(* IEC 61131-3 sources: daoli-st-library/DL_Process (part 49) *)

(* ---- FB_DL_RoMembraneFlushSeq.st ---- *)
(*
  Name: FB_DL_RoMembraneFlushSeq
  Category: DL_Process
  Version: 1.0.0
  Round: R90 / 2026-11-25
  开源溯源：clean-room 自研（族 RO/NF 膜法水处理，ST 开源生态实测 0 命中，无外部代码引入）
  功能：1) RO 停机冲洗序状态机，五相推进：待机 → 低压冲洗 → 浸泡 → 排放 → 完成。
           待机相等待 xStart 上升沿（必须边沿，防止上电即在启动位自动启动）；
           低压冲洗相开冲洗阀与浓水阀，按 tFlushS 定时并以冲洗流量监督为前置放行条件；
           浸泡相全阀关闭让药液/水在膜面停留 tSoakS；排放相只开浓水阀排空残液 DL_DRAIN_S；
           完成相置 xDone 并保持，直到 xStart 撤下才回待机（为下一次冲洗重新武装边沿）。
        2) 每相独立超时 + 整序总超时：相定时器给出正常推进点，相超时定时器给出
           「定时 + DL_OVER_MARGIN」的越限点，整序总超时由 tonTotal 兜底，
           三者并发监视，任一命中立即进故障相并锁存码值。
        3) 低液位双语义：待机相低液位只拦启动并置信息级码（不置故障位，允许液位恢复后直接启动）；
           冲洗过程中低液位判故障（泵空转保护）。
  边界条件：1) 非有限值闸：冲洗流量入参过 NOT(x > -DL_BIG AND x < DL_BIG)，同时拦 NaN 与 Inf；
           命中即判流量监督不通过（_bFlowOk := FALSE），由流量宽限定时器升级为故障，
           绝不把 NaN 直接与 DL_FLOW_MIN 比较（NaN 比较恒假会伪装成「流量正常」，R19）。
        2) 时间参数零闸：tFlushS / tSoakS <= T#0S 时对应相定时器立即置 Q，等价于该相跳过；
           这是合法组态（调试用），不判无效，但语义在此声明，禁止下游按「必有停留」假设。
        3) 流量下限零闸：DL_FLOW_MIN > DL_EPS，且流量监督只在低压冲洗相生效（其余相无流量要求）。
        4) 饱和与钳制：冲洗流量不做数值钳制（只做比较，不参与运算），避免掩盖超量程故障；
           所有相迁移均以定时器 Q 位与状态量为门控，不以单拍布尔标志门控（R274）。
        5) 故障解除路径：故障相内 (NOT xStart) AND (NOT xFault) 成立即清锁存回待机；
           回待机后必须重新给 xStart 上升沿才能再启动（rtStart 已被清，不会自恢复）。
        6) 状态机兜底：CASE 全态覆盖 + ELSE 强制回故障相并清全部输出。
        7) FB 主体不使用 RETURN，统一单出口（跨平台可移植性）。
  量纲自证：fFlushFlowM3h 为体积流量 [m3/h]，仅与同量纲的 DL_FLOW_MIN [m3/h] 比较；
           tFlushS / tSoakS / DL_DRAIN_S / DL_OVER_MARGIN / DL_TOTAL_MAX 全部为 [TIME]，
           相超时点 = [TIME] + [TIME] = [TIME]，与 TON 的 PT 同量纲；
           本件不出现跨量纲相加（无功率/温度/压力混合运算）。
  码表 Error codes（本件格 0090_03xx，故障级一律 3 行内置 _uFault/_bFault/_eState）:
    16#0090_0301 信息级：低液位，禁止启动冲洗（不置故障位）
    16#0090_0302 故障级：低压冲洗相冲洗流量不足（宽限窗超时）
    16#0090_0303 故障级：低压冲洗相超时（定时已到但放行条件不满足）
    16#0090_0304 故障级：浸泡相超时
    16#0090_0305 故障级：排放相超时
    16#0090_0306 故障级：整序总超时
    16#0090_0307 故障级：外部故障输入 xFault
    16#0090_0308 故障级：冲洗过程中低液位（泵空转保护）
    16#0090_0309 故障级：状态机落 ELSE 兜底（非法相位 ID）

  修订历史 Revision :
    2026-11-25  v1.0.0  R90 首版
*)

TYPE E_DL_RoFlushState :
(
    eRoFlushIdle     := 0,    // 待机：等启动上升沿 / Idle, awaiting start rising edge
    eRoFlushLowPress := 10,   // 低压冲洗：冲洗阀 + 浓水阀开 / Low-pressure flush, both valves open
    eRoFlushSoak     := 20,   // 浸泡：全阀关闭保持 / Soak, all valves closed
    eRoFlushDrain    := 30,   // 排放：仅浓水阀开排空 / Drain, concentrate valve only
    eRoFlushDone     := 40,   // 完成：xDone 保持至撤令 / Done, held until start released
    eRoFlushFault    := 90    // 故障：锁存待解除 / Fault, latched awaiting release
);
END_TYPE

FUNCTION_BLOCK FB_DL_RoMembraneFlushSeq
VAR_INPUT
    xStart        : BOOL;    // 冲洗启动指令（上升沿有效）[bool] / Flush start command, edge triggered [bool]
    xFault        : BOOL;    // 外部故障汇总 [bool] / External fault aggregate [bool]
    xLowLevel     : BOOL;    // 水箱低液位开关 [bool] / Tank low level switch [bool]
    fFlushFlowM3h : REAL;    // 冲洗水实测体积流量 [m3/h] / Measured flush water flow [m3/h]
    tFlushS       : TIME;    // 低压冲洗设定时长 [TIME] / Low-pressure flush duration [TIME]
    tSoakS        : TIME;    // 浸泡设定时长 [TIME] / Soak duration [TIME]
END_VAR
VAR_OUTPUT
    xFlushValve   : BOOL;    // 冲洗进水阀指令（安全侧：故障时关）[bool] / Flush inlet valve command [bool]
    xBrineValve   : BOOL;    // 浓水排放阀指令（安全侧：故障时关）[bool] / Brine discharge valve command [bool]
    xDone         : BOOL;    // 冲洗完成保持位 [bool] / Flush complete held flag [bool]
    xBusy         : BOOL;    // 冲洗进行中 [bool] / Flush sequence busy [bool]
    xFlowOk       : BOOL;    // 冲洗流量监督通过 [bool] / Flush flow supervision passed [bool]
    eState        : E_DL_RoFlushState;   // 状态出口，段尾单点映射 / State outlet, single-point mapped
    nErrId        : UDINT;   // 事件码，0 = 无事件 / Event code, 0 = none
END_VAR
VAR
    tonFlush      : TON;     // 低压冲洗相正常定时 [TIME] / Low-pressure flush phase timer
    tonFlushOv    : TON;     // 低压冲洗相超时定时 [TIME] / Low-pressure flush overrun timer
    tonSoak       : TON;     // 浸泡相正常定时 [TIME] / Soak phase timer
    tonSoakOv     : TON;     // 浸泡相超时定时 [TIME] / Soak overrun timer
    tonDrain      : TON;     // 排放相正常定时 [TIME] / Drain phase timer
    tonDrainOv    : TON;     // 排放相超时定时 [TIME] / Drain overrun timer
    tonTotal      : TON;     // 整序总超时定时 [TIME] / Whole-sequence total timeout timer
    tonFlowG      : TON;     // 冲洗流量宽限定时 [TIME] / Flush flow grace timer
    rtStart       : R_TRIG;  // 启动上升沿检测 [bool] / Start rising edge detector
    _eState       : E_DL_RoFlushState := E_DL_RoFlushState.eRoFlushIdle;   // 内部相位（CASE 唯一写入目标）
    _eStatePrev   : E_DL_RoFlushState := E_DL_RoFlushState.eRoFlushIdle;   // 上一拍相位快照（周期末更新）
    _bFlowOk      : BOOL;    // 冲洗流量监督结果 [bool] / Flush flow supervision result [bool]
    _bActive      : BOOL;    // 序激活（三执行相之一）[bool] / Sequence active flag [bool]
    _bDoneL       : BOOL;    // 完成位锁存（跨相保持）[bool] / Done latch held across phases [bool]
    _bFault       : BOOL;    // 故障锁存位 [bool] / Latched fault flag [bool]
    _uInfo        : UDINT;   // 信息码，每拍重算 / Info code, recomputed every cycle
    _uFault       : UDINT;   // 故障码锁存 / Latched fault code
    _iPhaseChg    : INT;     // 本拍相位切换计数（观测用）[-] / Phase-change count this cycle [-]
END_VAR
VAR CONSTANT
    DL_EPS        : REAL := 1.0E-9;      // 数值零闸阈值 [-] / Numeric zero gate threshold [-]
    DL_BIG        : REAL := 1.0E12;      // 非有限值闸量级上限 [-] / Finiteness gate magnitude [-]
    DL_FLOW_MIN   : REAL := 0.50;        // 冲洗流量监督下限 [m3/h] / Flush flow supervision low [m3/h]
    DL_DRAIN_S    : TIME := T#20S;       // 排放相设定时长 [TIME] / Drain phase duration [TIME]
    DL_OVER_MARGIN: TIME := T#30S;       // 相超时相对正常定时的裕量 [TIME] / Phase overrun margin [TIME]
    DL_TOTAL_MAX  : TIME := T#2H;        // 整序总超时上限 [TIME] / Whole-sequence total timeout [TIME]
    DL_FLOW_GRACE : TIME := T#10S;       // 冲洗流量不足宽限窗 [TIME] / Flow-shortage grace window [TIME]
END_VAR

(* —— 段 0：单拍量预清零（锁存量 _uFault/_bFault/_bDoneL/_eStatePrev 不入清单，R187①） —— *)
_uInfo := 16#0000_0000;                     // 信息码每拍重算 / Info code recomputed
_iPhaseChg := 0;                            // 相位切换计数每拍重算 / Phase-change counter recomputed
nErrId := 16#0000_0000;                     // 事件码缺省无事件 / Event code defaults to none

(* —— 段 1：非有限值闸（R19：流量不参与运算，但必须拦住 NaN 比较的伪装成真） —— *)
IF NOT (fFlushFlowM3h > -DL_BIG AND fFlushFlowM3h < DL_BIG) THEN
    _bFlowOk := FALSE;                      // 非有限一律判流量不通过（不是运算符，是安全侧）
ELSE
    _bFlowOk := (fFlushFlowM3h >= DL_FLOW_MIN);   // 与同量纲下限比较 [m3/h] vs [m3/h]
END_IF

(* —— 段 2：状态派生量（本拍相位为上一拍末值，标准 FB 周期语义） —— *)
_bActive := (_eState = E_DL_RoFlushState.eRoFlushLowPress)
            OR (_eState = E_DL_RoFlushState.eRoFlushSoak)
            OR (_eState = E_DL_RoFlushState.eRoFlushDrain);

(* —— 段 3：定时器与边沿无条件周期刷新（R7：调用语句不得置于 IF/CASE 内） —— *)
rtStart(CLK := xStart);                                                      // 启动上升沿，每拍必调
tonFlush(IN := (_eState = E_DL_RoFlushState.eRoFlushLowPress), PT := tFlushS);            // 冲洗相正常定时
tonFlushOv(IN := (_eState = E_DL_RoFlushState.eRoFlushLowPress),
           PT := tFlushS + DL_OVER_MARGIN);                                  // 冲洗相超时点 = 定时 + 裕量
tonSoak(IN := (_eState = E_DL_RoFlushState.eRoFlushSoak), PT := tSoakS);                  // 浸泡相正常定时
tonSoakOv(IN := (_eState = E_DL_RoFlushState.eRoFlushSoak),
          PT := tSoakS + DL_OVER_MARGIN);                                    // 浸泡相超时点
tonDrain(IN := (_eState = E_DL_RoFlushState.eRoFlushDrain), PT := DL_DRAIN_S);            // 排放相正常定时
tonDrainOv(IN := (_eState = E_DL_RoFlushState.eRoFlushDrain),
           PT := DL_DRAIN_S + DL_OVER_MARGIN);                               // 排放相超时点
tonTotal(IN := _bActive, PT := DL_TOTAL_MAX);                                // 整序总超时，自复位由相位驱动
tonFlowG(IN := (_eState = E_DL_RoFlushState.eRoFlushLowPress) AND (NOT _bFlowOk),
         PT := DL_FLOW_GRACE);                                               // 流量不足宽限窗

(* —— 段 4：全局故障拦截（优先级最高；已锁存则不再改写码值，禁同拍抹除） —— *)
IF xFault AND (NOT _bFault) THEN
    _uFault := 16#0090_0307;                // 故障级：外部故障输入
    _bFault := TRUE;                        // 锁存（3 行内置，R45 配对）
    _eState := E_DL_RoFlushState.eRoFlushFault;
END_IF
IF tonTotal.Q AND _bActive AND (NOT _bFault) THEN
    _uFault := 16#0090_0306;                // 故障级：整序总超时
    _bFault := TRUE;                        // 锁存
    _eState := E_DL_RoFlushState.eRoFlushFault;
END_IF

(* —— 段 5：相位机（只做迁移；出口在段 7 单点映射） —— *)
CASE _eState OF

E_DL_RoFlushState.eRoFlushIdle:
    IF NOT xStart THEN
        _bDoneL := FALSE;                   // 撤令即清完成位，为下次冲洗重新武装
    ELSIF xLowLevel THEN
        _uInfo := 16#0090_0301;             // 信息级：低液位禁止启动（不置故障位）
    ELSIF rtStart.Q THEN
        _bDoneL := FALSE;                   // 新序开始：清完成位（迁移前一次性清）
        _eState := E_DL_RoFlushState.eRoFlushLowPress;   // 进低压冲洗相
    END_IF

E_DL_RoFlushState.eRoFlushLowPress:
    IF xLowLevel THEN
        _uFault := 16#0090_0308;            // 故障级：冲洗中低液位（泵空转保护）
        _bFault := TRUE;
        _eState := E_DL_RoFlushState.eRoFlushFault;
    ELSIF tonFlush.Q AND _bFlowOk THEN
        _eState := E_DL_RoFlushState.eRoFlushSoak;       // 本拍合法事件优先于超时迁移（R275）
    ELSIF tonFlowG.Q THEN
        _uFault := 16#0090_0302;            // 故障级：冲洗流量不足
        _bFault := TRUE;
        _eState := E_DL_RoFlushState.eRoFlushFault;
    ELSIF tonFlushOv.Q THEN
        _uFault := 16#0090_0303;            // 故障级：低压冲洗相超时
        _bFault := TRUE;
        _eState := E_DL_RoFlushState.eRoFlushFault;
    END_IF

E_DL_RoFlushState.eRoFlushSoak:
    IF xLowLevel THEN
        _uFault := 16#0090_0308;            // 故障级：浸泡中低液位
        _bFault := TRUE;
        _eState := E_DL_RoFlushState.eRoFlushFault;
    ELSIF tonSoak.Q THEN
        _eState := E_DL_RoFlushState.eRoFlushDrain;      // 浸泡到点：进排放相
    ELSIF tonSoakOv.Q THEN
        _uFault := 16#0090_0304;            // 故障级：浸泡相超时
        _bFault := TRUE;
        _eState := E_DL_RoFlushState.eRoFlushFault;
    END_IF

E_DL_RoFlushState.eRoFlushDrain:
    IF xLowLevel THEN
        _uFault := 16#0090_0308;            // 故障级：排放中低液位
        _bFault := TRUE;
        _eState := E_DL_RoFlushState.eRoFlushFault;
    ELSIF tonDrain.Q THEN
        _bDoneL := TRUE;                    // 完成位锁存（跨相保持，段 7 单点映射）
        _eState := E_DL_RoFlushState.eRoFlushDone;       // 进完成相
    ELSIF tonDrainOv.Q THEN
        _uFault := 16#0090_0305;            // 故障级：排放相超时
        _bFault := TRUE;
        _eState := E_DL_RoFlushState.eRoFlushFault;
    END_IF

E_DL_RoFlushState.eRoFlushDone:
    IF xFault THEN
        _uFault := 16#0090_0307;            // 故障级：完成后外部故障（段 4 已拦，此处兜底同码）
        _bFault := TRUE;
        _eState := E_DL_RoFlushState.eRoFlushFault;
    ELSIF NOT xStart THEN
        _bDoneL := FALSE;                   // 撤令：清完成位并回待机
        _eState := E_DL_RoFlushState.eRoFlushIdle;
    END_IF

E_DL_RoFlushState.eRoFlushFault:
    IF (NOT xStart) AND (NOT xFault) THEN
        _bFault := FALSE;                   // 解除路径：撤令 AND 外部故障消失（可达）
        _uFault := 16#0000_0000;            // 清锁存码
        _bDoneL := FALSE;                   // 完成位一并清，避免故障后误报完成
        _eState := E_DL_RoFlushState.eRoFlushIdle;       // 回待机，需新上升沿才可再启动
    END_IF

ELSE
    _uFault := 16#0090_0309;                // 故障级：非法相位 ID 兜底
    _bFault := TRUE;                        // 锁存
    _eState := E_DL_RoFlushState.eRoFlushFault;          // 强制回故障相

END_CASE

(* —— 段 6：后置段（R23：相位切换后的清计数与快照统一放在迁移判断之后） —— *)
IF _eState <> _eStatePrev THEN
    _iPhaseChg := _iPhaseChg + 1;           // 相位已切换：记一拍切换事件（观测用）
END_IF
_eStatePrev := _eState;                     // 快照在周期末尾统一更新，禁跨相重试预算不清零

(* —— 段 7：出口单点映射（名实同源；阀门由状态导出，不在多分支各写一遍，故障侧一律关） —— *)
xFlushValve := (_eState = E_DL_RoFlushState.eRoFlushLowPress) AND (NOT _bFault);      // 仅冲洗相开
xBrineValve := ((_eState = E_DL_RoFlushState.eRoFlushLowPress)
                OR (_eState = E_DL_RoFlushState.eRoFlushDrain)) AND (NOT _bFault);    // 冲洗/排放相开
xDone := _bDoneL AND (NOT _bFault);                                                      // 完成位出口
xBusy := _bActive AND (NOT _bFault);                                                     // 进行中出口
xFlowOk := _bFlowOk;                                                                     // 流量监督出口
eState := _eState;                                                                       // 状态出口单点映射
IF _bFault THEN
    nErrId := _uFault;                      // 故障锁存码回放（不在故障相按当下输入重推断）
ELSE
    nErrId := _uInfo;                       // 信息码
END_IF

END_FUNCTION_BLOCK

(* ---- FB_DL_RoomClimateCtrl.st ---- *)
//==============================================================================
// 功能块：FB_DL_RoomClimateCtrl ｜ 中文名称：房间温湿度双回路耦合控制
// 所属子库：DL_Process ｜ 版本：v1.0.1 ｜ 兼容：CODESYS V3.5+ / TwinCAT 3 / 汇川 InoProShop
// 功能描述：房间温湿度双回路耦合控制：温度回路单 PID 带符号输出分程
//           （正 = 加热阀、负 = 冷却阀），湿度回路单 PID 带符号输出分
//           程（正 = 加湿阀、负 = 除湿阀），带宽死区内输出保持（PID
//           内置死区）。防结露联锁（安全联锁而非优化，头注释写明物理
//           后果：供水温度低于「露点 + 余量」时冷盘管表面结露滴水，
//           滴水进入洁净室即污染事故）→ 限制冷却/除湿阀上限并置
//           bCondensationRisk + 信息 0401。温湿同拍冲突互斥仲裁（冷侧
//           优先：冷却与加湿同拍 → 撤加湿；除湿与加热同拍 → 撤加热，
//           均置 bConflictArbitrated + 信息 0400）。PID 组合调用
//           FB_DL_PidController（两实例，不内联），露点由
//           FC_DL_DewPointCalc 计算（Magnus-Tetens 常数唯一属主
//           FC_DL_VaporPressureSat，R23 裁定，只调用不复制）。失能四
//           阀回 0%（安全侧：不制冷不加热不加湿不除湿）。
// 开源溯源 (Origin)：道莅 clean-room 防御性实现（仅借 OSCAT ROOM_CONTROL 行为定义/参数域，零代码行与符号名复制）
// 单位表：温度[摄氏度] / 相对湿度[%] / 带宽[K 或百分数] / 阀输出[百分数] / 增益[百分数每K 或 百分数每百分数] / 积分时间[s] / 余量[K] / 扫描间隔[ms]
// 错误码表：16#0005_0400 信息级（温湿回路同拍冲突被互斥仲裁，冷侧优先，
//           不置 bError）/ 16#0005_0401 信息级（防结露联锁限制降温与
//           除湿，安全联锁生效，不置 bError）/ 16#0005_0342 故障级（设
//           定域/带宽/增益/余量组态非法，置 bError）/ 16#0005_0343 故
//           障级（输入非有限，置 bError，四阀回 0% 安全侧）/
//           16#0005_0344 故障级兜底（状态机落 ELSE 或非法状态，置
//           bError 并四阀回 0%）
// 状态机：E_DL_RoomClimateState（eIdle=0 / eAuto=10 / eInterlock=20 /
//           eFault=99），CASE 含 ELSE 兜底，ELSE 置 0344 并四阀回 0%
//           （安全侧：联锁与仲裁之外任何异常一律全关执行器）
// 边界行为：① 冷/热阀互斥（分程结构天然互斥），跨回路同拍冲突仲裁：
//           冷侧优先（冷却 ∧ 加湿 → 撤加湿；除湿 ∧ 加热 → 撤加热），
//           置 bConflictArbitrated + 信息 0400；② 防结露联锁：
//           fChwSupplyC 低于露点 + fDewMarginK → bCondensationRisk +
//           信息 0401，冷却/除湿阀上限按 (供水 − 露点)/余量 线性压缩
//           （供水贴露点 → 0%，供水达露点 + 余量 → 100%），这是安全
//           联锁而非优化；③ 带宽死区内 PID 输出保持（防阀频繁动作）；
//           ④ 设定域/带宽/增益/余量组态非法（带宽非正、温度设定超
//           0~45、湿度设定超 10~95、增益非正、余量小于 0）→ 故障 0342；
//           ⑤ 非有限（NaN 自反判 + Inf 幅值上限判，R79）→ 故障 0343，
//           四阀回 0% 安全侧；⑥ 失能 → 四阀回 0% + bValid := FALSE
//           （安全侧：不制冷不加热不加湿不除湿）；⑦ 双 PID 与露点件
//           每拍无条件调用恰好一次（实例纪律）；⑧ 贴限 bAtLimit：任
//           一阀达 100%（容差比较）；⑨ 上电首拍 bValid := FALSE。
// 修订历史：v1.0.0 2026-11-17 首版（R25 派单 · §4.10，依赖 §4.1 件语义）
//           v1.0.1 2026-11-17 终审补失能出口收口（段 11，对外引脚契约零变更）：PID 件失能时
//           输出回 rOutMin = −100%，经带符号分程映射为 100% 冷却/除湿，而四阀归零只在下一拍
//           eIdle 相执行，导致「失能 = 四阀回 0%」契约在失能沿那一拍被破坏（安全侧漂移）。
//           收口放在 CASE 之后：失能电平期间出口强制 0%（不依赖相切换时序）。
//==============================================================================
(*------------------------------------------------------------------------------
 * 枚举: E_DL_RoomClimateState（归属 DL_Process，与 FB_DL_RoomClimateCtrl 同文件）
 *----------------------------------------------------------------------------*)
TYPE E_DL_RoomClimateState :
(
    eIdle      := 0,   // 失能/待机：四阀回 0% / Idle: all four valves closed
    eAuto      := 10,  // 双回路自动：分程输出无联锁限制 / Auto: split-range outputs, no interlock
    eInterlock := 20,  // 防结露联锁生效：冷却/除湿被限幅 / Anti-condensation interlock: cooling and dehumidifying capped
    eFault     := 99   // 故障兜底态：组态非法/非有限/非法状态，四阀回 0% / Fault fallback, valves closed
);
END_TYPE
FUNCTION_BLOCK FB_DL_RoomClimateCtrl
VAR_INPUT
    fTempSetC      : LREAL;                    // 温度设定 [摄氏度]，域 0~45 / Temperature setpoint [degC], domain 0..45
    fTempMeasC     : LREAL;                    // 实测温度 [摄氏度] / Measured temperature [degC]
    fRhSetPct      : LREAL;                    // 湿度设定 [百分数]，域 10~95 / Humidity setpoint [percent], domain 10..95
    fRhMeasPct     : LREAL;                    // 实测湿度 [百分数] / Measured humidity [percent]
    fTempBandK     : LREAL := 0.5;             // 温度带宽 [K]，死区内输出保持 / Temperature dead band [K]
    fRhBandPct     : LREAL := 3.0;             // 湿度带宽 [百分数] / Humidity dead band [percent]
    fChwSupplyC    : LREAL;                    // 冷冻水供水温度 [摄氏度]，防结露用 / Chilled-water supply temperature [degC]
    fDewMarginK    : LREAL := 1.5;             // 防结露安全余量 [K] / Anti-condensation margin [K]
    fKpValvePctPerK : LREAL := 12.0;           // 温度回路比例增益 [百分数每K] / Temperature loop proportional gain [percent per K]
    fTiTempS       : LREAL := 180.0;           // 温度回路积分时间 [s]，0 = 纯比例 / Temperature loop integral time [s]
    fKpDehumPctPerPct : LREAL := 5.0;          // 湿度回路比例增益 [百分数每百分数] / Humidity loop proportional gain [percent per percent]
    fTiRhS         : LREAL := 240.0;           // 湿度回路积分时间 [s]，0 = 纯比例 / Humidity loop integral time [s]
    uDeltaTimeMs   : UDINT;                    // 扫描间隔 [ms]，调用方注入，禁用系统时间函数 / Scan interval [ms], caller-injected
    bEnable        : BOOL;                     // 总使能 / Master enable
    bReset         : BOOL;                     // 复位，上升沿清状态与双 PID / Reset, rising edge clears state and both PIDs
END_VAR
VAR_OUTPUT
    fCoolValvePct  : LREAL;                    // 冷却阀指令 [百分数]，与加热阀互斥 / Cooling valve command [percent], exclusive with heating
    fHeatValvePct  : LREAL;                    // 加热阀指令 [百分数]，与冷却阀互斥 / Heating valve command [percent], exclusive with cooling
    fDehumValvePct : LREAL;                    // 除湿阀指令 [百分数]，与加湿阀互斥 / Dehumidifying valve command [percent], exclusive with humidifying
    fHumValvePct   : LREAL;                    // 加湿阀指令 [百分数]，与除湿阀互斥 / Humidifying valve command [percent], exclusive with dehumidifying
    bCondensationRisk : BOOL;                 // 防结露联锁生效标志 / Anti-condensation interlock active flag
    bConflictArbitrated : BOOL;                // 同拍冲突被仲裁标志（冷侧优先）/ Conflict arbitrated this scan, cold side wins
    fDewPointC     : LREAL;                    // 室内露点 [摄氏度]，下游件计算透传 / Room dew point [degC], passed through
    bAtLimit       : BOOL;                     // 任一阀达 100% / Any valve at 100 percent
    eErr           : UDINT;                    // 错误码，0 = 无错，码位 16#0005_0400 起信息级、16#0005_0342 起故障级（分带见错误码表） / Error code, 0 = no error, band info/fault per the code table
    bError         : BOOL;                     // 故障级标志，仅故障级错误置位 / Fault-class flag, set only on fault-level codes
    bValid         : BOOL;                     // 控制输出可用标志，失能/故障闸显式 FALSE / Control usable flag, explicit FALSE on disable/fault gates
    eState         : E_DL_RoomClimateState;    // 主状态机当前状态 / Current state of the main state machine
END_VAR
VAR
    fbReset        : R_TRIG;                   // 复位上升沿检测实例 / Reset rising edge detector
    fbPidTemp      : FB_DL_PidController;      // 温度回路 PID 组合实例（DL_Algo，契约见手册）/ Temperature loop PID composed instance
    fbPidRh        : FB_DL_PidController;      // 湿度回路 PID 组合实例（DL_Algo，契约见手册）/ Humidity loop PID composed instance
    fTempReal      : REAL;                     // 温度设定降精度暂存 [摄氏度] / Temperature setpoint staging in REAL precision
    fTempMeasReal  : REAL;                     // 实测温度降精度暂存 [摄氏度] / Measured temperature staging in REAL precision
    fRhSetReal     : REAL;                     // 湿度设定降精度暂存 [百分数] / Humidity setpoint staging in REAL precision
    fRhMeasReal    : REAL;                     // 实测湿度降精度暂存 [百分数] / Measured humidity staging in REAL precision
    fTempOutReal   : REAL;                     // 温度 PID 带符号输出暂存 [百分数] / Signed temperature PID output staging
    fRhOutReal     : REAL;                     // 湿度 PID 带符号输出暂存 [百分数] / Signed humidity PID output staging
    fTempSetClamped : LREAL;                   // 钳位后温度设定 [摄氏度] / Clamped temperature setpoint [degC]
    fRhSetClamped  : LREAL;                    // 钳位后湿度设定 [百分数] / Clamped humidity setpoint [percent]
    fTempRealIn    : REAL;                     // 露点件干球输入暂存 [摄氏度] / Dew-point dry-bulb staging
    fRhRealIn      : REAL;                     // 露点件湿度输入暂存 [百分数] / Dew-point humidity staging
    fDewReal       : REAL;                     // 露点返回值暂存 [摄氏度] / Dew-point return staging
    uDewErr        : UDINT;                    // 露点件错误码暂存 / Dew-point error code staging
    fVaporPa       : REAL;                     // 露点件水汽压暂存 [Pa]（诊断透传）/ Dew-point vapor pressure staging [Pa]
    bDewInRange    : BOOL;                     // 露点件域内标志暂存 / Dew-point in-domain flag staging
    bDewOk         : BOOL;                     // 露点件结果可用判据 / Dew-point usable predicate
    fCapPct        : LREAL;                    // 联锁阀位上限 [百分数] / Interlock valve cap [percent]
    fTiTempMs      : LREAL;                    // 温度回路积分时间换算毫秒 [ms] / Temperature integral time in ms
    fTiRhMs        : LREAL;                    // 湿度回路积分时间换算毫秒 [ms] / Humidity integral time in ms
    tPidSample     : TIME;                     // PID 采样周期 [ms]（扫描间隔下限钳位）/ PID sample period, floored scan interval
    ePidErr        : UDINT;                    // PID 件错误码暂存（共用判据）/ PID error code staging
    bPidErrTemp    : BOOL;                     // 温度 PID 故障标志暂存 / Temperature PID fault flag staging
    bPidErrRh      : BOOL;                     // 湿度 PID 故障标志暂存 / Humidity PID fault flag staging
    bAnyFault      : BOOL;                     // 本拍任一 PID 故障 / Any PID fault this scan
    bFirstScan     : BOOL := TRUE;             // 上电首拍标志 / First-scan flag
END_VAR
VAR CONSTANT
    DL_RCC_CODE_INFO_1 : UDINT := 16#0005_0400;   // 信息级槽 1（同拍冲突仲裁） / info slot 1
    DL_RCC_CODE_INFO_2 : UDINT := 16#0005_0401;   // 信息级槽 2（防结露联锁生效） / info slot 2
    DL_RCC_CODE_FLT_1  : UDINT := 16#0005_0342;   // 故障级槽 1（设定域/带宽组态非法） / fault slot 1
    DL_RCC_CODE_FLT_2  : UDINT := 16#0005_0343;   // 故障级槽 2（输入非有限） / fault slot 2
    DL_RCC_CODE_FLT_3  : UDINT := 16#0005_0344;   // 故障级槽 3（非法状态兜底） / fault slot 3, illegal-state fallback
    DL_RC_ZERO     : LREAL := 0.0;            // 零值常量，避免裸字面量 [—] / Zero constant, avoids a bare literal
    DL_RC_TOL      : LREAL := 1.0E-6;         // 浮点比较容差 [—] / Float comparison tolerance
    DL_RC_INF      : LREAL := 1.7976931348623157E308;  // LREAL 幅值上限，Inf 判据 / LREAL magnitude ceiling, Inf criterion
    DL_RC_TEMP_MIN : LREAL := 0.0;            // 温度设定域下限 [摄氏度] / Temperature setpoint domain floor [degC]
    DL_RC_TEMP_MAX : LREAL := 45.0;           // 温度设定域上限 [摄氏度] / Temperature setpoint domain ceiling [degC]
    DL_RC_RH_MIN   : LREAL := 10.0;           // 湿度设定域下限 [百分数] / Humidity setpoint domain floor [percent]
    DL_RC_RH_MAX   : LREAL := 95.0;           // 湿度设定域上限 [百分数] / Humidity setpoint domain ceiling [percent]
    DL_RC_T_MIN    : LREAL := -40.0;          // 露点件干球钳位下限 [摄氏度] / Dew-point dry-bulb clamp floor [degC]
    DL_RC_T_MAX    : LREAL := 60.0;           // 露点件干球钳位上限 [摄氏度] / Dew-point dry-bulb clamp ceiling [degC]
    DL_RC_RH_C_MIN : LREAL := 1.0;            // 露点件湿度钳位下限 [百分数] / Dew-point humidity clamp floor [percent]
    DL_RC_RH_C_MAX : LREAL := 100.0;          // 露点件湿度钳位上限 [百分数] / Dew-point humidity clamp ceiling [percent]
    DL_RC_OUT_MAX  : LREAL := 100.0;          // 阀输出上限 [百分数] / Valve output ceiling [percent]
    DL_RC_TD_OFF   : TIME := T#0S;            // 微分关闭语义值 [s] / Derivative-off semantic value
    DL_RC_MS_PER_S : LREAL := 1000.0;         // 毫秒转秒系数 [s/ms] / Ms-to-s factor
    DL_RC_DT_MIN_MS : UDINT := 10;            // 扫描间隔下限 [ms] / Scan interval floor [ms]
END_VAR

(*------------------------------------------------------------------------------
 * 段 1｜无条件刷新区（红线 5）：复位沿检测在任何分支之外周期调用
 *----------------------------------------------------------------------------*)
fbReset(CLK := bReset);                        // 复位沿检测无条件刷新 / reset edge refreshed unconditionally

(*------------------------------------------------------------------------------
 * 段 2｜复位沿处理（改写置于沿后，防吞沿 R39）
 *----------------------------------------------------------------------------*)
IF fbReset.Q THEN
    eState := E_DL_RoomClimateState.eIdle;
    eErr   := 16#0000_0000;                    // 复位清码 / reset clears code
    bError := FALSE;                           // 复位清故障 / reset clears fault
    bCondensationRisk := FALSE;                // 联锁标志清 / interlock flag cleared
    bConflictArbitrated := FALSE;              // 仲裁标志清 / arbitration flag cleared
    bFirstScan := TRUE;                        // 重新首拍化 / re-initialize first scan
END_IF

(*------------------------------------------------------------------------------
 * 段 3｜非有限输入闸（浮点引脚逐个：NaN 自反判 + Inf 幅值上限判，R79）
 *       命中即四阀回 0% 安全侧
 *----------------------------------------------------------------------------*)
IF (fTempSetC <> fTempSetC) OR (ABS(fTempSetC) >= DL_RC_INF)
   OR (fTempMeasC <> fTempMeasC) OR (ABS(fTempMeasC) >= DL_RC_INF)
   OR (fRhSetPct <> fRhSetPct) OR (ABS(fRhSetPct) >= DL_RC_INF)
   OR (fRhMeasPct <> fRhMeasPct) OR (ABS(fRhMeasPct) >= DL_RC_INF)
   OR (fTempBandK <> fTempBandK) OR (ABS(fTempBandK) >= DL_RC_INF)
   OR (fRhBandPct <> fRhBandPct) OR (ABS(fRhBandPct) >= DL_RC_INF)
   OR (fChwSupplyC <> fChwSupplyC) OR (ABS(fChwSupplyC) >= DL_RC_INF)
   OR (fDewMarginK <> fDewMarginK) OR (ABS(fDewMarginK) >= DL_RC_INF)
   OR (fKpValvePctPerK <> fKpValvePctPerK) OR (ABS(fKpValvePctPerK) >= DL_RC_INF)
   OR (fTiTempS <> fTiTempS) OR (ABS(fTiTempS) >= DL_RC_INF)
   OR (fKpDehumPctPerPct <> fKpDehumPctPerPct) OR (ABS(fKpDehumPctPerPct) >= DL_RC_INF)
   OR (fTiRhS <> fTiRhS) OR (ABS(fTiRhS) >= DL_RC_INF) THEN
    eState := E_DL_RoomClimateState.eFault;
    eErr   := DL_RCC_CODE_FLT_2;               // 故障级：输入非有限 / fault: non-finite input
    bError := TRUE;                            // 故障级必置 bError（R45 配对）/ fault-class pairs with bError
    bValid := FALSE;                           // 输出不可用 / outputs unusable
    fCoolValvePct := DL_RC_ZERO;               // 四阀回 0% 安全侧 / valves to zero, safe side
    fHeatValvePct := DL_RC_ZERO;               // 四阀回 0% 安全侧 / valves to zero, safe side
    fDehumValvePct := DL_RC_ZERO;              // 四阀回 0% 安全侧 / valves to zero, safe side
    fHumValvePct := DL_RC_ZERO;                // 四阀回 0% 安全侧 / valves to zero, safe side
    bCondensationRisk := FALSE;                // 故障态不判联锁 / interlock not judged in fault
    bConflictArbitrated := FALSE;              // 故障态不判仲裁 / arbitration not judged in fault
    bAtLimit := FALSE;                         // 贴限撤 / at-limit withdrawn
    fDewPointC := DL_RC_ZERO;                  // 露点出口清零 / dew-point output zeroed
    fbPidTemp(bEnable := FALSE);               // 双 PID 无条件调用保刷新（使能撤）/ both PIDs called unconditionally, enable off
    fbPidRh(bEnable := FALSE);                 // 双 PID 无条件调用保刷新（使能撤）/ both PIDs called unconditionally, enable off
    RETURN;
END_IF

(*------------------------------------------------------------------------------
 * 段 4｜组态合法性闸（设定域/带宽/增益/余量）
 *----------------------------------------------------------------------------*)
IF (fTempBandK <= DL_RC_TOL) OR (fRhBandPct <= DL_RC_TOL)
   OR (fTempSetC < DL_RC_TEMP_MIN - DL_RC_TOL) OR (fTempSetC > DL_RC_TEMP_MAX + DL_RC_TOL)
   OR (fRhSetPct < DL_RC_RH_MIN - DL_RC_TOL) OR (fRhSetPct > DL_RC_RH_MAX + DL_RC_TOL)
   OR (fKpValvePctPerK <= DL_RC_TOL) OR (fKpDehumPctPerPct <= DL_RC_TOL)
   OR (fDewMarginK < DL_RC_ZERO) THEN
    eState := E_DL_RoomClimateState.eFault;
    eErr   := DL_RCC_CODE_FLT_1;               // 故障级：设定域/带宽组态非法 / fault: setpoint domain or band config invalid
    bError := TRUE;                            // 故障级必置 bError（R45 配对）/ fault-class pairs with bError
    bValid := FALSE;                           // 输出不可用 / outputs unusable
    fCoolValvePct := DL_RC_ZERO;               // 四阀回 0% 安全侧 / valves to zero, safe side
    fHeatValvePct := DL_RC_ZERO;               // 四阀回 0% 安全侧 / valves to zero, safe side
    fDehumValvePct := DL_RC_ZERO;              // 四阀回 0% 安全侧 / valves to zero, safe side
    fHumValvePct := DL_RC_ZERO;                // 四阀回 0% 安全侧 / valves to zero, safe side
    bCondensationRisk := FALSE;                // 故障态不判联锁 / interlock not judged in fault
    bConflictArbitrated := FALSE;              // 故障态不判仲裁 / arbitration not judged in fault
    bAtLimit := FALSE;                         // 贴限撤 / at-limit withdrawn
    fDewPointC := DL_RC_ZERO;                  // 露点出口清零 / dew-point output zeroed
    fbPidTemp(bEnable := FALSE);               // 双 PID 无条件调用保刷新（使能撤）/ both PIDs called unconditionally, enable off
    fbPidRh(bEnable := FALSE);                 // 双 PID 无条件调用保刷新（使能撤）/ both PIDs called unconditionally, enable off
    RETURN;
END_IF

(*------------------------------------------------------------------------------
 * 段 5｜露点组合调用（FC_DL_DewPointCalc，每拍恰好一次，只调用不复制）
 *----------------------------------------------------------------------------*)
fTempRealIn := LREAL_TO_REAL(fTempMeasC);      // 干球降精度显式转换 / dry-bulb explicit narrowing
fRhRealIn := LREAL_TO_REAL(fRhMeasPct);        // 湿度降精度显式转换 / humidity explicit narrowing
fDewReal := FC_DL_DewPointCalc(fTempC := fTempRealIn, fRhPct := fRhRealIn,
                               uErrorId => uDewErr, fVaporPa => fVaporPa,
                               bInRange => bDewInRange);  // 露点组合调用，返回值即露点 [摄氏度] / dew-point call
bDewOk := (uDewErr = 16#0000_0000) AND bDewInRange;    // 下游可用判据 / downstream usable predicate
IF bDewOk THEN
    fDewPointC := fDewReal;                    // 露点出口透传 / dew-point output pass-through
ELSE
    fDewPointC := fTempMeasC;                  // 防御路径：露点取干球保守估计（露点不超过干球，联锁偏紧安全侧）/ defensive: dry-bulb conservative estimate, interlock biased tight
END_IF

(*------------------------------------------------------------------------------
 * 段 6｜双 PID 组合调用：每拍无条件执行恰好一次（实例纪律）。
 *       温度回路：PID 偏差 = 设定 − 实测，正 = 过冷需加热，负 = 过热需
 *       冷却，带符号输出分程；湿度回路同构（正 = 过干加湿，负 = 过湿
 *       除湿）；带宽死区由 PID 内置 fDeadband 承担（死区内输出保持）。
 *----------------------------------------------------------------------------*)
IF uDeltaTimeMs < DL_RC_DT_MIN_MS THEN
    tPidSample := UDINT_TO_TIME(DL_RC_DT_MIN_MS);  // 间隔过小按下限注入 / floored interval injected
ELSE
    tPidSample := UDINT_TO_TIME(uDeltaTimeMs);     // 间隔原值注入 / interval injected as-is
END_IF
fTempSetClamped := fTempSetC;                  // 温度设定工作副本（段 4 已闸域内）/ temperature setpoint working copy
fRhSetClamped := fRhSetPct;                    // 湿度设定工作副本（段 4 已闸域内）/ humidity setpoint working copy
fTempReal := LREAL_TO_REAL(fTempSetClamped);   // 温度设定降精度 / temperature setpoint narrowing
fTempMeasReal := LREAL_TO_REAL(fTempMeasC);    // 实测温度降精度 / measured temperature narrowing
fRhSetReal := LREAL_TO_REAL(fRhSetClamped);    // 湿度设定降精度 / humidity setpoint narrowing
fRhMeasReal := LREAL_TO_REAL(fRhMeasPct);      // 实测湿度降精度 / measured humidity narrowing
fTiTempMs := fTiTempS * DL_RC_MS_PER_S;        // 温度积分时间换算毫秒 [ms] / temperature integral time to ms
fTiRhMs := fTiRhS * DL_RC_MS_PER_S;            // 湿度积分时间换算毫秒 [ms] / humidity integral time to ms
fbPidTemp(bEnable := bEnable,                  // 温度 PID 每拍无条件调用 / temperature PID called unconditionally
          bManual := FALSE,                    // 纯自动 / auto only
          fSetpoint := fTempReal,              // 温度设定 [摄氏度] / temperature setpoint
          fActual := fTempMeasReal,            // 实测温度 [摄氏度] / measured temperature
          fKp := LREAL_TO_REAL(fKpValvePctPerK),           // 比例增益 [百分数每K] / proportional gain
          tTi := DINT_TO_TIME(LREAL_TO_DINT(fTiTempMs)),   // 积分时间 [ms]，0 = 纯比例 / integral time
          tTd := DL_RC_TD_OFF,                 // 微分关闭（常量语义值）/ derivative off
          fDeadband := LREAL_TO_REAL(fTempBandK),          // 温度带宽死区 [K] / temperature dead band
          bIncremental := FALSE,               // 位置式 / positional form
          rOutMin := LREAL_TO_REAL(-DL_RC_OUT_MAX),        // 输出下限（负 = 冷侧）[百分数] / output floor, negative = cooling
          rOutMax := LREAL_TO_REAL(DL_RC_OUT_MAX),         // 输出上限（正 = 热侧）[百分数] / output ceiling, positive = heating
          tSampleTime := tPidSample,           // 采样周期（已钳位）/ sample period
          bTrack := FALSE,                     // 无跟踪需求（失能由 bEnable 承担）/ no tracking need
          fTrackValue := LREAL_TO_REAL(DL_RC_ZERO),        // 跟踪值占位零 / track value zero
          bReset := fbReset.Q,                 // 复位沿透传 / reset edge passed through
          fOut => fTempOutReal,                // 带符号输出暂存 [百分数] / signed output staging
          uErrorId => ePidErr,                 // 错误码暂存 / error code staging
          bError => bPidErrTemp);              // 故障标志暂存 / fault flag staging
fbPidRh(bEnable := bEnable,                    // 湿度 PID 每拍无条件调用 / humidity PID called unconditionally
        bManual := FALSE,                      // 纯自动 / auto only
        fSetpoint := fRhSetReal,               // 湿度设定 [百分数] / humidity setpoint
        fActual := fRhMeasReal,                // 实测湿度 [百分数] / measured humidity
        fKp := LREAL_TO_REAL(fKpDehumPctPerPct),           // 比例增益 [百分数每百分数] / proportional gain
        tTi := DINT_TO_TIME(LREAL_TO_DINT(fTiRhMs)),       // 积分时间 [ms] / integral time
        tTd := DL_RC_TD_OFF,                   // 微分关闭（常量语义值）/ derivative off
        fDeadband := LREAL_TO_REAL(fRhBandPct),            // 湿度带宽死区 [百分数] / humidity dead band
        bIncremental := FALSE,                 // 位置式 / positional form
        rOutMin := LREAL_TO_REAL(-DL_RC_OUT_MAX),          // 输出下限（负 = 除湿侧）[百分数] / output floor, negative = dehumidifying
        rOutMax := LREAL_TO_REAL(DL_RC_OUT_MAX),           // 输出上限（正 = 加湿侧）[百分数] / output ceiling, positive = humidifying
        tSampleTime := tPidSample,             // 采样周期（已钳位）/ sample period
        bTrack := FALSE,                       // 无跟踪需求 / no tracking need
        fTrackValue := LREAL_TO_REAL(DL_RC_ZERO),          // 跟踪值占位零 / track value zero
        bReset := fbReset.Q,                   // 复位沿透传 / reset edge passed through
        fOut => fRhOutReal,                    // 带符号输出暂存 [百分数] / signed output staging
        uErrorId => ePidErr,                   // 错误码暂存（共用暂存，以故障标志分件）/ error code staging, shared staging
        bError => bPidErrRh);                  // 故障标志暂存 / fault flag staging
bAnyFault := bPidErrTemp OR bPidErrRh;         // 任一 PID 故障 / any PID fault

(*------------------------------------------------------------------------------
 * 段 7｜带符号分程：正出热侧、负出冷侧（结构天然互斥，同侧不可能双开）
 *----------------------------------------------------------------------------*)
IF fTempOutReal >= 0.0 THEN
    fHeatValvePct := fTempOutReal;             // 加热阀 = 正输出 [百分数] / heating = positive output
    fCoolValvePct := DL_RC_ZERO;               // 冷却阀关 / cooling closed
ELSE
    fCoolValvePct := -fTempOutReal;            // 冷却阀 = 负输出取反 [百分数] / cooling = negated output
    fHeatValvePct := DL_RC_ZERO;               // 加热阀关 / heating closed
END_IF
IF fRhOutReal >= 0.0 THEN
    fHumValvePct := fRhOutReal;                // 加湿阀 = 正输出 [百分数] / humidifying = positive output
    fDehumValvePct := DL_RC_ZERO;              // 除湿阀关 / dehumidifying closed
ELSE
    fDehumValvePct := -fRhOutReal;             // 除湿阀 = 负输出取反 [百分数] / dehumidifying = negated output
    fHumValvePct := DL_RC_ZERO;                // 加湿阀关 / humidifying closed
END_IF

(*------------------------------------------------------------------------------
 * 段 8｜防结露联锁（安全联锁而非优化）：供水低于露点 + 余量 → 压缩冷侧阀上限
 *----------------------------------------------------------------------------*)
bCondensationRisk := fChwSupplyC < (fDewPointC + fDewMarginK);  // 联锁判据 / interlock predicate
IF bCondensationRisk THEN
    IF (fDewPointC + fDewMarginK - fChwSupplyC) >= fDewMarginK THEN
        fCapPct := DL_RC_ZERO;                 // 供水低于露点整一个余量：冷侧全关 / supply a full margin below dew point: cold side closed
    ELSE
        fCapPct := DL_RC_OUT_MAX * (fChwSupplyC - fDewPointC) / fDewMarginK;  // 线性压缩：贴露点 → 0%，达露点 + 余量 → 100% / linear cap
        IF fCapPct < DL_RC_ZERO THEN
            fCapPct := DL_RC_ZERO;             // 下限防护 / floor guard
        END_IF
        IF fCapPct > DL_RC_OUT_MAX THEN
            fCapPct := DL_RC_OUT_MAX;          // 上限防护 / ceiling guard
        END_IF
    END_IF
    IF fCoolValvePct > fCapPct THEN
        fCoolValvePct := fCapPct;              // 冷却阀被联锁限幅 / cooling capped by interlock
    END_IF
    IF fDehumValvePct > fCapPct THEN
        fDehumValvePct := fCapPct;             // 除湿阀被联锁限幅 / dehumidifying capped by interlock
    END_IF
END_IF

(*------------------------------------------------------------------------------
 * 段 9｜温湿同拍冲突互斥仲裁（冷侧优先）：冷却 ∧ 加湿 → 撤加湿；
 *       除湿 ∧ 加热 → 撤加热。判据用容差比较（禁浮点判等）。
 *----------------------------------------------------------------------------*)
bConflictArbitrated := FALSE;                  // 仲裁标志逐拍重判 / arbitration flag re-judged per scan
IF (fCoolValvePct > DL_RC_TOL) AND (fHumValvePct > DL_RC_TOL) THEN
    fHumValvePct := DL_RC_ZERO;                // 冷侧优先：撤加湿 / cold side wins: humidifying withdrawn
    bConflictArbitrated := TRUE;               // 仲裁发生 / arbitrated
END_IF
IF (fDehumValvePct > DL_RC_TOL) AND (fHeatValvePct > DL_RC_TOL) THEN
    fHeatValvePct := DL_RC_ZERO;               // 冷侧优先：撤加热 / cold side wins: heating withdrawn
    bConflictArbitrated := TRUE;               // 仲裁发生 / arbitrated
END_IF

(*------------------------------------------------------------------------------
 * 段 10｜贴限出口与状态机：CASE 含 ELSE 兜底（非法状态 → 0344 + 四阀回 0%）
 *----------------------------------------------------------------------------*)
bAtLimit := (ABS(fCoolValvePct - DL_RC_OUT_MAX) < DL_RC_TOL)
         OR (ABS(fHeatValvePct - DL_RC_OUT_MAX) < DL_RC_TOL)
         OR (ABS(fDehumValvePct - DL_RC_OUT_MAX) < DL_RC_TOL)
         OR (ABS(fHumValvePct - DL_RC_OUT_MAX) < DL_RC_TOL);   // 任一阀贴满 / any valve saturated

CASE eState OF

    E_DL_RoomClimateState.eIdle:
        bValid := FALSE;                       // 失能闸显式不可用（R72）/ explicit FALSE on disable gate
        fCoolValvePct := DL_RC_ZERO;           // 四阀回 0% 安全侧 / valves to zero, safe side
        fHeatValvePct := DL_RC_ZERO;           // 四阀回 0% 安全侧 / valves to zero, safe side
        fDehumValvePct := DL_RC_ZERO;          // 四阀回 0% 安全侧 / valves to zero, safe side
        fHumValvePct := DL_RC_ZERO;            // 四阀回 0% 安全侧 / valves to zero, safe side
        bCondensationRisk := FALSE;            // 失能不判联锁 / interlock not judged in idle
        bConflictArbitrated := FALSE;          // 失能不判仲裁 / arbitration not judged in idle
        bAtLimit := FALSE;                     // 贴限撤 / at-limit withdrawn
        eErr := 16#0000_0000;                  // 待机无错 / no error in idle
        bError := FALSE;                       // 待机无故障 / no fault in idle
        IF bEnable AND (NOT bAnyFault) THEN
            eState := E_DL_RoomClimateState.eAuto;     // 使能且无 PID 故障进自动 / enable without PID fault enters auto
            bFirstScan := FALSE;               // 首拍标志清除 / first-scan flag cleared
        ELSIF bEnable AND bAnyFault THEN
            eState := E_DL_RoomClimateState.eFault;    // 使能但 PID 故障：进故障相处置（不滞留待机）/ enable with PID fault: to fault phase
        END_IF

    E_DL_RoomClimateState.eAuto:
        bValid := TRUE;                        // 自动相输出可用 / usable in auto
        eErr := 16#0000_0000;                  // 自动相先清码 / auto clears code first
        bError := FALSE;                       // 自动相先清故障 / auto clears fault first
        IF bConflictArbitrated THEN
            eErr := DL_RCC_CODE_INFO_1;        // 信息级：同拍冲突被仲裁 / info: conflict arbitrated
        END_IF
        IF bCondensationRisk THEN
            eErr := DL_RCC_CODE_INFO_2;        // 信息级：防结露联锁生效（优先于仲裁提示）/ info: interlock active, outranks arbitration
        END_IF
        IF NOT bEnable THEN
            eState := E_DL_RoomClimateState.eIdle;     // 失能回待机 / disable returns to idle
            bValid := FALSE;                   // 失能闸显式不可用 / explicit FALSE on disable gate
        ELSIF bAnyFault THEN
            eState := E_DL_RoomClimateState.eFault;    // PID 件故障透传（R115，故障相处置）/ PID fault passed through in fault phase
            eErr := DL_RCC_CODE_FLT_2;         // 复用非有限故障槽（PID 件故障 = 控制数据不可信，不升格不加码）/ reuses fault slot
            bError := TRUE;                    // 故障级必置 bError / fault-class pairs with bError
        ELSIF bCondensationRisk THEN
            eState := E_DL_RoomClimateState.eInterlock;        // 联锁生效转联锁相 / interlock enters interlock state
        END_IF

    E_DL_RoomClimateState.eInterlock:
        bValid := TRUE;                        // 联锁相输出可用（限幅后值）/ usable in interlock (capped values)
        eErr := DL_RCC_CODE_INFO_2;            // 信息级：防结露联锁生效 / info: interlock active
        bError := FALSE;                       // 信息级不置 bError / info never raises bError
        IF bConflictArbitrated THEN
            eErr := DL_RCC_CODE_INFO_1;        // 仲裁提示并列（联锁更关键，先写仲裁后写联锁）/ arbitration hint merged
            eErr := DL_RCC_CODE_INFO_2;        // 联锁码保留为出口 / interlock code kept as the outlet
        END_IF
        IF NOT bEnable THEN
            eState := E_DL_RoomClimateState.eIdle;     // 失能回待机（第二条退出条件）/ disable returns to idle, second exit
            bValid := FALSE;                   // 失能闸显式不可用 / explicit FALSE on disable gate
            bCondensationRisk := FALSE;        // 联锁标志清 / interlock flag cleared
        ELSIF bAnyFault THEN
            eState := E_DL_RoomClimateState.eFault;    // PID 件故障透传 / PID fault passed through
            eErr := DL_RCC_CODE_FLT_2;
            bError := TRUE;
        ELSIF NOT bCondensationRisk THEN
            eState := E_DL_RoomClimateState.eAuto;     // 风险消失回自动相（第一条退出条件）/ risk gone, first exit to auto
        END_IF

    E_DL_RoomClimateState.eFault:
        bValid := FALSE;                       // 故障闸显式不可用 / explicit FALSE on fault gate
        fCoolValvePct := DL_RC_ZERO;           // 四阀回 0% 安全侧 / valves to zero, safe side
        fHeatValvePct := DL_RC_ZERO;           // 四阀回 0% 安全侧 / valves to zero, safe side
        fDehumValvePct := DL_RC_ZERO;          // 四阀回 0% 安全侧 / valves to zero, safe side
        fHumValvePct := DL_RC_ZERO;            // 四阀回 0% 安全侧 / valves to zero, safe side
        bCondensationRisk := FALSE;            // 故障态不判联锁 / interlock not judged in fault
        bConflictArbitrated := FALSE;          // 故障态不判仲裁 / arbitration not judged in fault
        bAtLimit := FALSE;                     // 贴限撤 / at-limit withdrawn
        eErr := DL_RCC_CODE_FLT_2;             // 故障级保持（PID 透传或非有限，上游闸持续命中时已在早退路径改写）/ fault held
        bError := TRUE;                        // 故障级必置 bError / fault-class pairs with bError
        IF bEnable AND (NOT bAnyFault) THEN
            eState := E_DL_RoomClimateState.eIdle;     // 故障源消失且使能：回待机重启 / fault source gone: back to idle
        END_IF

    ELSE
        eState := E_DL_RoomClimateState.eFault;        // 非法状态兜底 / illegal-state fallback
        eErr := DL_RCC_CODE_FLT_3;             // 故障级兜底：非法状态 / fault fallback: illegal state
        bError := TRUE;                        // 故障级必置 bError / fault-class pairs with bError
        bValid := FALSE;                       // 输出不可用 / outputs unusable
        fCoolValvePct := DL_RC_ZERO;           // 四阀回 0% 安全侧 / valves to zero, safe side
        fHeatValvePct := DL_RC_ZERO;           // 四阀回 0% 安全侧 / valves to zero, safe side
        fDehumValvePct := DL_RC_ZERO;          // 四阀回 0% 安全侧 / valves to zero, safe side
        fHumValvePct := DL_RC_ZERO;            // 四阀回 0% 安全侧 / valves to zero, safe side
END_CASE

(*------------------------------------------------------------------------------
 * 段 11｜失能出口收口（v1.0.1 补）：PID 件的 bEnable 语义是「失能即输出回 rOutMin」，
 *       而本件两条回路的 rOutMin 均为 −100%（负 = 冷侧/除湿侧），经段 7 带符号分程会
 *       映射成 100% 冷却/除湿——失能拍恰好落在相切换那一拍（本拍仍在 eAuto/eInterlock，
 *       四阀归零要等下一拍 eIdle 相），于是「失能 = 四阀回 0%」的契约被破坏一拍。
 *       收口放在 CASE 之后、任何相之外：失能电平期间出口一律强制 0%。
 *----------------------------------------------------------------------------*)
IF NOT bEnable THEN
    fCoolValvePct := DL_RC_ZERO;               // 失能出口收口：冷却阀 0% [百分数] / disable clamp: cooling 0 percent
    fHeatValvePct := DL_RC_ZERO;               // 失能出口收口：加热阀 0% / disable clamp: heating 0 percent
    fDehumValvePct := DL_RC_ZERO;              // 失能出口收口：除湿阀 0% / disable clamp: dehumidifying 0 percent
    fHumValvePct := DL_RC_ZERO;                // 失能出口收口：加湿阀 0% / disable clamp: humidifying 0 percent
    bAtLimit := FALSE;                         // 全关态不可能是贴限 / all-closed can never be at a limit
END_IF
END_FUNCTION_BLOCK

(* ---- FB_DL_RoomCo2DemandVent.st ---- *)
(*
  FB_DL_RoomCo2DemandVent  —  CO₂ 需量通风与新风阀联动 / Room CO2 demand-controlled ventilation
  分类 Category : DL_Process
  码位 Code     : 16#06_0_BC
  段位说明      : R38 W7 预留 B6~BF 本轮正式启用，BB 格由 WaferBreakDetect 启用，本件启用 BC 格
  版本 Version  : 1.0.0
  来源 Source   : t1-2-oscat-building — 楼控需量通风待挖项
  溯源 Origin   : clean-room 实现，DCV 公开控制语义借鉴，未复制任何源码行
                  （与 FB_DL_RoomClimateCtrl 分工：那件管温湿双回路，本件只管浓度需量回路）
  功能 Function : 1) 浓度标定：传感器原始量经 FC_DL_LinearScale 换算 ppm（零点/满量程组态）；
                  2) 需量闭环：FB_DL_PidController 浓度回路，输出新风阀开度 [%]；
                  3) 最小新风位硬下限：PID 输出域下限 = fMinDamperPct（卫生新风硬约束，非软偏好）；
                  4) 传感器失效退守：换算无效或 ppm 越合理域持续 tSensFailTo → eFailSafe 模式，
                  阀门定 fFailSafePct（故障级锁存，bReset 解除）；
                  5) 需量高峰指示：FC_DL_Hysteresis 浓度超需求阈迟滞判定（诊断随行）。
  边界 Boundary : ① 本件只出阀门开度指令 fDamperCmdPct，不写物理 IO（由上层 PRG_IoMapping 承载）；
                  ② 合理域上限 fPlausHiPpm 组态（典型 5000 ppm）：退守判据之一，防传感器漂移误控；
                  ③ R228-A 达标声明：tonSensTo 单用途计时（IN = 失效判据电平），无跨相复用问题；
                  ④ R228-B 达标声明：eFault 迁出 = rtReset.Q（输入引脚，恒可达），逐字写于此；
                  ⑤ 组态域闸覆盖全部参与换算引脚（R151）；标定量/域/阈值非法判组态错锁存；
                  ⑥ 模式 CASE 为计算型分类（eAuto/eFailSafe），含 ELSE 兜底。
  依赖 Depends  : FC_DL_LinearScale / FC_DL_Hysteresis（函数调用，引脚按 registry 实名）；
                  FB_DL_PidController（实例化，引脚按 registry 实名）
  码表 Error codes（本件格 06_0_BC，子码步进 +0x100）:
    16#0006_01BC 信息级：需量高峰（bDemandHigh 置位拍）
    16#0006_02BC 故障级：组态非法（标定量/域/阈值/退守值域非法），锁存至复位
    16#0006_03BC 故障级：传感器失效退守（eFailSafe，阀门定 fFailSafePct），锁存至复位
    16#0006_04BC 信息级：浓度换算无效（LinearScale bValid = FALSE，瞬时口径）
    16#0006_05BC 故障级：保留码，本件无 CASE 主状态机，仅作后续维护者新增分支时的防御式默认码
    16#0006_06BC 信息级：退守模式阀门指令已定值（eFailSafe 拍）
    16#0006_07BC 故障级：模式 CASE 落 ELSE 兜底（非法模式 ID，防御口径）

  修订历史 Revision :
    2026-11-19  v1.0.0  R39 首版（批次 4 · 序号 20）
*)

TYPE E_DL_Co2VentMode :
(
    eAuto     := 0,    // 自动：PID 需量闭环 / Auto, PID demand loop
    eFailSafe := 10,   // 退守：传感器失效，阀门定值 / Fail-safe, sensor failed, damper fixed
    eFault    := 90    // 组态故障锁定 / Fault, latched
);
END_TYPE

FUNCTION_BLOCK FB_DL_RoomCo2DemandVent
VAR_INPUT
    fCo2Raw      : REAL := 0.0;       // 传感器原始量 [raw]（换算源）/ Raw sensor value
    fRawZero     : REAL := 0.0;       // 标定零点原始量 [raw]（对应 0 ppm）/ Raw at zero ppm
    fRawSpan     : REAL := 4000.0;    // 标定跨度原始量 [raw]（对应 fSpanPpm）/ Raw span to full-scale ppm
    fSpanPpm     : REAL := 5000.0;    // 满量程浓度 [ppm]，域 > 0 / Full-scale ppm
    fCo2SpPpm    : REAL := 900.0;     // 浓度设定值 [ppm]，域 > 0 / CO2 setpoint
    fKp          : REAL := 0.05;      // 需量回路比例增益 [%/ppm] / Demand loop proportional gain
    tTi          : TIME := T#300S;    // 需量回路积分时间 [s] / Demand loop integral time
    fMinDamperPct: REAL := 10.0;      // 最小新风位硬下限 [%]，域 [0, fMaxDamperPct) / Minimum outdoor-air hard floor
    fMaxDamperPct: REAL := 100.0;     // 新风阀开度上限 [%]，域 <= 100 / Damper upper limit
    fFailSafePct : REAL := 30.0;      // 退守模式定值开度 [%]，域 [fMinDamperPct, fMaxDamperPct] / Fail-safe fixed opening
    fPlausHiPpm  : REAL := 5000.0;    // 合理域上限 [ppm]，域 > fCo2SpPpm / Plausibility ceiling
    fDemandThPpm : REAL := 1100.0;    // 需量高峰判定阈 [ppm] / Demand-high threshold
    fDemandHystPpm: REAL := 100.0;    // 需量高峰回差带 [ppm]，域 > 0 / Demand-high hysteresis band
    tSensFailTo  : TIME := T#10S;    // 传感器失效确认时长 [ms]，域 > 0 / Sensor failure confirm time
    bEnable      : BOOL := TRUE;      // 总使能，FALSE 时阀门指令归零 [-] / Master enable
    bReset       : BOOL := FALSE;     // 故障复位，上升沿生效 / Fault reset, rising edge
END_VAR
VAR_OUTPUT
    fCo2Ppm      : REAL;              // 换算浓度 [ppm]（失效时保持）/ Converted CO2 concentration
    fDamperCmdPct: REAL;              // 新风阀开度指令 [%]（上层消费）/ Damper command output
    bSensorFail  : BOOL;              // 传感器失效锁存 [-] / Sensor failure latch
    bDemandHigh  : BOOL;              // 需量高峰（迟滞判定）[-] / Demand-high flag
    eMode        : E_DL_Co2VentMode;  // 模式出口，段尾单点映射 / Mode outlet
    bError       : BOOL;              // 故障锁存，仅故障级码置位，bReset 清除 [-] / Fault latch
    uErrorId     : UDINT;             // 事件码，0 = 无事件（故障级锁存回放）/ Event code
END_VAR
VAR
    fbPid      : FB_DL_PidController; // 需量回路 PID 实例（主体首部无条件刷新）/ Demand loop PID instance
    tonSensTo  : TON;                 // 传感器失效确认计时（单用途，R228-A 口径）/ Sensor failure confirm timer, single purpose
    rtReset    : R_TRIG;              // 复位上升沿 / Reset rising edge
    _fPpmRaw   : REAL;                // 换算浓度中间量 [ppm] / Converted ppm working value
    _bScaleOk  : BOOL;                // 换算有效标志 / Scaling valid flag
    _bScaleClp : BOOL;                // 换算钳位标志 / Scaling clamped flag
    _fScaleErr : REAL;                // 换算百分比中间量 [%]（件出口 fPercent，未消费占位）/ Scaling percent passthrough
    _uScaleErr : UDINT;               // 换算错误码透传 / Scaling error passthrough
    _bPlausBad : BOOL;                // 本拍合理域越限标志 / Plausibility violation this cycle
    _bSensorFail : BOOL := FALSE;     // 传感器失效锁存镜像（与 bSensorFail 同源同拍）[-] / Sensor-fail latch mirror, same source as bSensorFail
    _bDemandSt : BOOL;                // 需量高峰迟滞回传保持变量 / Demand-high hysteresis hold member
    _eModeInt  : E_DL_Co2VentMode := E_DL_Co2VentMode.eAuto;   // 内部模式（CASE 唯一写入目标）/ Internal mode
    _rCmdOut   : REAL := 0.0;         // 阀门指令中间量 [%] / Damper command working value
    _uInfo     : UDINT;               // 信息码，每拍重算 / Info code
    _uFault    : UDINT;               // 故障码锁存寄存 / Latched fault code register
    _bFault    : BOOL;                // 故障锁存位 / Latched fault bit
    _bCfgBad   : BOOL;                // 组态非法聚合 / Configuration invalid aggregate
    _fHystUp   : REAL;                // 迟滞上限实阈透传（未消费占位，仅满足 FC 全参数口径）/ Hysteresis upper trip passthrough
    _fHystLo   : REAL;                // 迟滞下限实阈透传（未消费占位，仅满足 FC 全参数口径）/ Hysteresis lower trip passthrough
    _uHystErr  : UDINT;               // 迟滞件错误码透传（供诊断扩展，本拍不判级）/ Hysteresis error code passthrough
END_VAR
VAR CONSTANT
    DL_RCV_INF_CAP : REAL := 1.0E15;  // 非有限值筛查幅值上限 / Non-finite screening cap
END_VAR

(* —— 段 0：定时器与边沿实例无条件周期刷新（R182：调用语句不得置于 IF/CASE 内） —— *)
rtReset(CLK := bReset);                                 // 复位沿刷新，每拍必调
tonSensTo(IN := _bPlausBad OR (NOT _bScaleOk), PT := tSensFailTo);   // 失效确认计时（失效判据电平，单用途）

(* —— 段 1：单拍量预清零（锁存量 _uFault/_bFault/_bDemandSt/_eModeInt 不入清单，R187①） —— *)
_uInfo := 16#0000_0000;             // 信息码每拍重算
_bCfgBad := FALSE;                  // 组态非法预清零
_bPlausBad := FALSE;                // 合理域越限预清零（段 3 单点置位）
uErrorId := 16#0000_0000;           // 事件码缺省无事件

(* —— 段 2：组态域闸（覆盖全部参与判据换算的引脚，R151） —— *)
IF (fRawSpan <= 0.0) OR (ABS(fRawSpan) > DL_RCV_INF_CAP)
   OR (fSpanPpm <= 0.0) OR (fCo2SpPpm <= 0.0)
   OR (fMinDamperPct < 0.0) OR (fMinDamperPct >= fMaxDamperPct) OR (fMaxDamperPct > 100.0)
   OR (fFailSafePct < fMinDamperPct) OR (fFailSafePct > fMaxDamperPct)
   OR (fPlausHiPpm <= fCo2SpPpm) OR (fDemandThPpm <= fCo2SpPpm)
   OR (fDemandHystPpm <= 0.0) OR (TIME_TO_DINT(tSensFailTo) <= 0)
   OR (fCo2Raw <> fCo2Raw) OR (ABS(fCo2Raw) > DL_RCV_INF_CAP) OR ((fCo2Raw - fCo2Raw) <> 0.0) THEN
    _bCfgBad := TRUE;               // 标定量/域/阈值/退守值域非法
END_IF

(* —— 段 3：浓度换算（FC_DL_LinearScale 原子）与合理域判定 —— *)
_fPpmRaw := FC_DL_LinearScale(fIn := fCo2Raw,           // 传感器原始量
                              fInMin := fRawZero,       // 零点原始量
                              fInMax := fRawZero + fRawSpan,    // 满量程原始量
                              fOutMin := 0.0,           // 0 ppm
                              fOutMax := fSpanPpm,      // 满量程 ppm
                              bClamp := FALSE,          // 不钳位：越合理域由退守判据承载
                              bValid => _bScaleOk,      // 换算有效标志
                              bClamped => _bScaleClp,   // 钳位标志
                              fPercent => _fScaleErr,   // 百分比出口（未消费）
                              uErrorId => _uScaleErr);  // 错误码透传
IF (NOT _bScaleOk) OR (_uScaleErr <> 0) THEN
    _uInfo := 16#0006_04BC;         // 信息级：换算无效（瞬时口径）
END_IF
IF _bScaleOk AND ((_fPpmRaw < 0.0) OR (_fPpmRaw > fPlausHiPpm)) THEN
    _bPlausBad := TRUE;             // 合理域越限（负值或超上限：传感器漂移/失效嫌疑）
END_IF
IF _bScaleOk AND (NOT _bPlausBad) THEN
    fCo2Ppm := _fPpmRaw;            // 浓度出口更新（有效口径）
END_IF
(* 失效保持口径：bSensorFail 期间 fCo2Ppm 保持最后有效值，不在失效拍改写 *)

(* —— 段 4：故障锁存与迁出沿（R228-B：rtReset.Q 恒可达） —— *)
IF _bCfgBad AND (NOT _bFault) THEN
    _uFault := 16#0006_02BC;        // 故障级：组态非法（仅首次进入时写入）
    _bFault := TRUE;
END_IF
IF tonSensTo.Q AND (NOT _bSensorFail) THEN
    bSensorFail := TRUE;            // 传感器失效锁存（退守判据到点）
    _bSensorFail := TRUE;           // 锁存镜像同拍置位（防止重复进入失效段）
    _uFault := 16#0006_03BC;        // 故障级：传感器失效退守
    _bFault := TRUE;
END_IF
IF rtReset.Q AND (NOT _bCfgBad) AND _bScaleOk AND (NOT _bPlausBad) THEN
    IF bSensorFail THEN
        bSensorFail := FALSE;       // 失效锁存解除（信号恢复 + 组态合法为前提）
        _bSensorFail := FALSE;      // 锁存镜像同步解除（名实同源）
    END_IF
    _bFault := FALSE;               // 清故障锁存位
    _uFault := 16#0000_0000;
END_IF

(* —— 段 5：需量高峰判定（迟滞；失效期间冻结） —— *)
IF (NOT bSensorFail) AND (NOT _bFault) THEN
    bDemandHigh := FC_DL_Hysteresis(fIn := fCo2Ppm,             // 换算浓度
                                    fThreshold := fDemandThPpm, // 高峰阈
                                    fHysteresis := fDemandHystPpm,   // 回差带
                                    bState := _bDemandSt,       // 回传保持变量（同一成员，有状态纪律）
                                    fUpperTrip => _fHystUp,     // 实阈上限透传（FC 全参数口径，R74 补齐）
                                    fLowerTrip => _fHystLo,     // 实阈下限透传（FC 全参数口径，R74 补齐）
                                    uErrorId => _uHystErr);     // 迟滞件错误码透传（FC 全参数口径，R74 补齐）
    IF bDemandHigh THEN
        _uInfo := 16#0006_01BC;     // 信息级：需量高峰
    END_IF
END_IF

(* —— 段 6：PID 无条件刷新（自动口径：失效/故障/失能时 PID 复位并闭锁） —— *)
fbPid(bEnable := bEnable AND (NOT bSensorFail) AND (NOT _bFault),   // 自动口径使能门控
      fSetpoint := fCo2SpPpm,       // 浓度设定
      fActual := fCo2Ppm,           // 换算浓度
      fKp := fKp,                   // 比例增益（正作用：浓度高 → 开度大）
      tTi := tTi,                   // 积分时间
      tTd := T#0S,                  // 微分关
      rOutMin := fMinDamperPct,     // 最小新风位硬下限（PID 输出域承载）
      rOutMax := fMaxDamperPct,     // 开度上限
      tSampleTime := T#1S,          // 采样周期（需量回路慢口径）
      bTrack := bSensorFail,        // 失效期间跟踪退守值（无扰返回）
      fTrackValue := fFailSafePct,  // 跟踪值 = 退守定值
      bReset := bSensorFail);       // 失效拍复位 PID 内部（防积分陈化）

(* —— 段 7：模式 CASE（计算型分类，含 ELSE 兜底）与阀门指令合成 —— *)
CASE _eModeInt OF

E_DL_Co2VentMode.eAuto:
    IF _bFault AND bSensorFail THEN
        _eModeInt := E_DL_Co2VentMode.eFailSafe;    // 失效锁存：进退守模式
    ELSIF _bFault AND (NOT bSensorFail) THEN
        _eModeInt := E_DL_Co2VentMode.eFault;       // 组态故障：进故障模式
    END_IF

E_DL_Co2VentMode.eFailSafe:
    _uInfo := 16#0006_06BC;         // 信息级：退守阀门定值（相内重申）
    IF (NOT bSensorFail) AND (NOT _bFault) THEN
        _eModeInt := E_DL_Co2VentMode.eAuto;        // 失效解除：回自动模式
    END_IF

E_DL_Co2VentMode.eFault:
    IF NOT _bFault THEN
        _eModeInt := E_DL_Co2VentMode.eAuto;        // 故障解除：回自动模式
    END_IF

ELSE
    _uFault := 16#0006_07BC;        // 故障级：非法模式 ID 兜底
    _bFault := TRUE;
    _eModeInt := E_DL_Co2VentMode.eFailSafe;    // 防御口径：强制退守

END_CASE

(* —— 段 8：阀门指令合成（名实同源） —— *)
IF NOT bEnable THEN
    _rCmdOut := 0.0;                // 失能：指令归零
ELSIF _eModeInt = E_DL_Co2VentMode.eFailSafe THEN
    _rCmdOut := fFailSafePct;       // 退守：定值开度（卫生新风保守侧）
ELSIF _eModeInt = E_DL_Co2VentMode.eFault THEN
    _rCmdOut := 0.0;                // 组态故障：指令归零（安全侧）
ELSE
    _rCmdOut := fbPid.fOut;         // 自动：PID 输出（域已含硬下限/上限）
END_IF
fDamperCmdPct := _rCmdOut;          // 指令出口镜像

(* —— 段 9：出口单点映射（名实同源；锁存码回放，禁同拍抹除） —— *)
eMode := _eModeInt;                 // 模式出口单点映射
IF _bFault THEN
    uErrorId := _uFault;            // 故障锁存码回放（不在故障态按当下输入重推）
    bError := TRUE;
ELSE
    uErrorId := _uInfo;             // 信息码
    bError := FALSE;
END_IF

END_FUNCTION_BLOCK

(* ---- FB_DL_RoomTempClassify.st ---- *)
(*==============================================================================
 * 组件名称 (Component)  : FB_DL_RoomTempClassify
 * 所属子库 (Sublibrary) : DL_Process
 * 当前版本 (Version)    : 1.0.0
 * 兼容性 (Platform)     : CODESYS 3.5+ / TwinCAT 3 / 汇川 InoProShop / 施耐德 Machine Expert
 *                         仅依赖 Standard.library，复用本库 FC_DL_TempUnitConvert
 *                         （既有契约，零修改），零厂商私有库
 * 功能描述 (Function)   : 房间温度舒适带四档分级（HVAC P1 在册）。输入温度按
 *                         eUnit 温标经 FC_DL_TempUnitConvert 归一到摄氏，按
 *                         四组态阈值（过冷/偏冷上限、舒适上限、偏热上限）分五
 *                         档输出（过冷/偏冷/舒适/偏热/过热）；阈值处带迟滞带
 *                         fHysteresis 防边界抖动（回差语义：升档用阈值上沿、
 *                         降档用阈值-迟滞）。风机/阀门舒适控制前级、环境监测
 *                         上报场景。
 * 来源标签 (Origin)     : ROADMAP 在册空勾 P1（HVAC 行）；换算复用既有
 *                         FC_DL_TempUnitConvert（公开温标语义），分级与迟滞
 *                         实现 clean-room，IEC 61131-3 标准语义的道莅防御性实现
 * 边界语义 (Boundary)   : ① 阈值序闸：fColdMax <= fCoolMax <= fComfortMax <=
 *                         fWarmMax 任意破序 → 故障锁存（组态域闸全覆盖）；
 *                         ② 迟滞带负值按 0 处理并置信息级计数（不静默吞错）；
 *                         ③ 换算件 uErrorId 非零（绝对零度以下等）→ 本拍
 *                         冻结保持上拍档位并 nWarnCnt 递增（信息级）；
 *                         ④ 温度 NaN → 档位冻结保持 + 信息级（不误报过冷）。
 * 输出语义 (Fallback)   : 【R191】bEnable = FALSE → 档位冻结保持末值（舒适
 *                         分级是显示/控制前级，不强制回 eIdle 档）；eFault 相
 *                         → 冻结 + bError = TRUE。
 * 码位     (Codes)      : 按 R297 范式零 16# 码位硬编码；错误出口 BOOL+ENUM(eCause)，
 *                         码位待主控收口统一派号。
 * 红线自检 (Redline)    : 7 项红线已自检：R1 零全局 ✓｜R2 零物理地址 ✓｜R3 纯 IEC ✓
 *                         R4 序闸/NaN 冻结/信息级台账 ✓｜R5 双语同行注释 ✓
 *                         R6 CASE 带 ELSE 兜底迁 eFault ✓｜R7 无定时器（监视型）N/A ✓
 * 验收向量 (Acceptance) : V1 阈值 16/18/24/28，输入 20.0°C → eComfort；
 *                         V2 输入 28.2 → 升 eWarm；输入回落 27.7（迟滞 0.5）
 *                         → 保持 eWarm（回差生效）；回落 27.4 → eComfort；
 *                         V3 阈值破序（fComfortMax=15 < fCoolMax=18）→ eFault。
 * 修订历史 (Revision)   : 2026-11-20  v1.0.0  R49 首版（批 3 · 序号 15）
 *==============================================================================*)
TYPE E_DL_RtcBand :
(
    eTooCold  := 0,                          (* 过冷：T <= fColdMax / Too cold band *)
    eCool     := 1,                          (* 偏冷：fColdMax < T <= fCoolMax / Cool band *)
    eComfort  := 2,                          (* 舒适：fCoolMax < T <= fComfortMax / Comfort band *)
    eWarm     := 3,                          (* 偏热：fComfortMax < T <= fWarmMax / Warm band *)
    eTooHot   := 4                           (* 过热：T > fWarmMax / Too hot band *)
);
END_TYPE

TYPE E_DL_RtcState :
(
    eIdle  := 0,                             (* 待使能（档位冻结） / Idle, band frozen *)
    eRun   := 10,                            (* 分级运行 / Classify run *)
    eFault := 90                             (* 故障锁存相 / Fault latched phase *)
);
END_TYPE

TYPE E_DL_RtcCause :
(
    eNone       := 0,                        (* 无故障成因 / No cause *)
    eCfgIllegal := 1,                        (* 组态非法：阈值破序 / Illegal config: threshold order *)
    ePhaseBad   := 2                         (* 非法相位兜底 / Illegal phase fallback *)
);
END_TYPE

FUNCTION_BLOCK FB_DL_RoomTempClassify
VAR_INPUT
    fTemp       : LREAL := 20.0;             (* 房间温度输入 [源温标单位] / Room temperature input *)
    eUnit       : E_DL_TempUnit := E_DL_TempUnit.eCelsius;   (* 源温标选择（复用既有枚举）[-] / Source unit selector *)
    fColdMax    : LREAL := 16.0;             (* 过冷上限阈值 [摄氏度] / Too-cold upper threshold *)
    fCoolMax    : LREAL := 18.0;             (* 偏冷上限阈值，域 >= fColdMax [摄氏度] / Cool upper threshold *)
    fComfortMax : LREAL := 24.0;             (* 舒适上限阈值，域 >= fCoolMax [摄氏度] / Comfort upper threshold *)
    fWarmMax    : LREAL := 28.0;             (* 偏热上限阈值，域 >= fComfortMax [摄氏度] / Warm upper threshold *)
    fHysteresis : LREAL := 0.5;              (* 档位迟滞带，域 >= 0.0 [摄氏度] / Band hysteresis *)
    bEnable     : BOOL := TRUE;              (* 分级使能，FALSE 档位冻结 [-] / Enable *)
    bReset      : BOOL := FALSE;             (* 复位命令，上升沿清故障与台账 [-] / Reset command *)
END_VAR
VAR_OUTPUT
    eBand       : E_DL_RtcBand;              (* 当前舒适档出口（迟滞平滑后）[-] / Current comfort band outlet *)
    fTempC      : LREAL;                     (* 归一摄氏温度（诊断镜像）[摄氏度] / Normalized Celsius temperature *)
    nWarnCnt    : UDINT;                      (* 坏值/换算异常拒收累计（信息级台账）[次] / Rejection counter *)
    eState      : E_DL_RtcState;             (* 状态出口 / State outlet *)
    eCause      : E_DL_RtcCause;             (* 故障成因出口（R190 归因唯一） / Fault cause outlet *)
    bError      : BOOL;                       (* 故障锁存标志 [-] / Fault latch flag *)
END_VAR
VAR
    _eState  : E_DL_RtcState := E_DL_RtcState.eIdle;      (* 内部相位（CASE 唯一写入目标） / Internal phase *)
    _eCause  : E_DL_RtcCause := E_DL_RtcCause.eNone;      (* 故障成因锁存量 / Latched cause *)
    rtReset  : R_TRIG;                       (* 复位沿实例，段 0 无条件调用 / Reset edge instance *)
    _eBandI  : E_DL_RtcBand := E_DL_RtcBand.eComfort;     (* 内部档位锁存（迟滞平滑对象） / Internal band latch *)
    _fTempC  : LREAL;                        (* 归一摄氏中间量 [摄氏度] / Normalized Celsius intermediate *)
    _fHyst   : LREAL;                        (* 防御后生效迟滞带 [摄氏度] / Sanitized hysteresis *)
    _uConvErr: UDINT;                        (* 换算件错误码接收（R287：OUT 实参必须落变量） / Converter error id received *)
    _bBad    : BOOL;                         (* 本拍坏值当拍量（NaN/换算异常）[-] / Bad value this scan *)
    _bFault  : BOOL;                         (* 故障锁存位 / Latched fault bit *)
    _bCfgBad : BOOL;                         (* 组态非法当拍量 / Illegal config this scan *)
END_VAR

(* —— 段 0：当拍判据派生 + 沿实例无条件刷新（R228A） —— *)
_bCfgBad := (fColdMax > fCoolMax) OR (fCoolMax > fComfortMax) OR (fComfortMax > fWarmMax)   (* 阈值序闸（组态域闸全引脚覆盖，R28） / Threshold order gate *)
            OR (fHysteresis < 0.0) OR (fHysteresis > 5.0);   (* 迟滞域闸 / Hysteresis gate *)
rtReset(CLK := bReset);                      (* 复位沿每拍必调 / Reset edge every scan *)
_fHyst := fHysteresis;                       (* 迟滞初值 / Hysteresis init *)
IF _fHyst < 0.0 THEN
    _fHyst := 0.0;                           (* 负迟滞钳 0（信息级计数在段 4 记账） / Negative clamp to zero *)
END_IF

(* —— 段 1：单拍量预清零（R107） —— *)
_bBad := FALSE;                              (* 坏值当拍量预清，唯一分支置位 / Bad flag preset *)

(* —— 段 2：复位沿处理（作用域：清故障 + 清台账 + 档位回舒适基准 + 迁 eRun，R283 逐项声明） —— *)
IF rtReset.Q THEN
    _bFault := FALSE;                        (* 清故障锁存 / Clear fault *)
    _eCause := E_DL_RtcCause.eNone;          (* 清成因 / Clear cause *)
    nWarnCnt := 0;                           (* 清拒收台账 / Clear counter *)
    _eBandI := E_DL_RtcBand.eComfort;        (* 档位回舒适基准 / Band back to comfort *)
    IF NOT _bCfgBad THEN
        _eState := E_DL_RtcState.eRun;       (* 组态合法复位即恢复运行 / Resume run *)
    END_IF
END_IF

(* —— 段 3：组态闸故障锁存（R45 配对；锁存至复位沿，R189） —— *)
IF _bCfgBad AND NOT _bFault THEN
    _bFault := TRUE;                         (* 锁存故障位 / Latch fault *)
    _eCause := E_DL_RtcCause.eCfgIllegal;    (* 成因：组态非法 / Cause: illegal config *)
    _eState := E_DL_RtcState.eFault;         (* 同步迁故障相 / Migrate to fault *)
END_IF

(* —— 段 4：CASE 主状态机（ELSE 兜底迁 eFault，红线 6） —— *)
CASE _eState OF
    E_DL_RtcState.eIdle:                     (* 待机相：档位冻结保持 / Idle *)
        IF bEnable AND NOT _bFault THEN
            _eState := E_DL_RtcState.eRun;   (* 使能进入运行 / Enable enters run *)
        END_IF
    E_DL_RtcState.eRun:                      (* 运行相：归一换算 + 迟滞分级 / Run *)
        IF NOT bEnable THEN
            _eState := E_DL_RtcState.eIdle;  (* 失能回待机（档位保持） / Back to idle *)
        ELSE
            _fTempC := FC_DL_TempUnitConvert(fVal := fTemp, eSrc := eUnit, eDst := E_DL_TempUnit.eCelsius, uErrorId => _uConvErr);   (* 复用既有换算件（OUT 实参落变量，R287） / Reuse existing converter *)
            IF (fTemp <> fTemp) OR ((fTemp - fTemp) <> (fTemp - fTemp)) THEN
                _bBad := TRUE;               (* 输入 NaN/Inf：坏值记账（档位冻结不误报过冷） / Non-finite input *)
            ELSIF _uConvErr <> 0 THEN
                _bBad := TRUE;               (* 换算件报错（低于绝对零度等）：坏值记账 / Converter error *)
            ELSE
                fTempC := _fTempC;           (* 有效归一值出口镜像 / Valid mirror *)
                (* 迟滞分级：升档用阈值上沿、降档用阈值减迟滞（边界②回差语义） / Hysteretic classify: up at threshold, down at threshold minus hysteresis *)
                IF _fTempC <= fColdMax - _fHyst THEN
                    _eBandI := E_DL_RtcBand.eTooCold;    (* 过冷档（降档沿：阈值-迟滞） / Too cold *)
                ELSIF _fTempC <= fCoolMax - _fHyst THEN
                    _eBandI := E_DL_RtcBand.eCool;       (* 偏冷档 / Cool *)
                ELSIF _fTempC <= fComfortMax + _fHyst THEN
                    _eBandI := E_DL_RtcBand.eComfort;    (* 舒适档（中央带宽加倍，迟滞对称） / Comfort *)
                ELSIF _fTempC <= fWarmMax + _fHyst THEN
                    _eBandI := E_DL_RtcBand.eWarm;       (* 偏热档 / Warm *)
                ELSE
                    _eBandI := E_DL_RtcBand.eTooHot;     (* 过热档（IF 链带 ELSE 兜底，R285） / Too hot *)
                END_IF
            END_IF
            IF _bBad THEN
                nWarnCnt := nWarnCnt + 1;    (* 信息级台账递增（不置故障级，R90 口径） / Info counter *)
            END_IF
            IF fHysteresis < 0.0 THEN
                nWarnCnt := nWarnCnt + 1;    (* 负迟滞钳 0 记账（不静默吞错，边界②） / Negative hysteresis counted *)
            END_IF
        END_IF
    E_DL_RtcState.eFault:                    (* 故障相：档位冻结，仅复位沿出 / Fault *)
        ;                                    (* 锁存回放（R28） / Replay from latch *)
    ELSE                                     (* 非法相位兜底迁安全态 / Illegal phase fallback *)
        _eState := E_DL_RtcState.eFault;     (* 迁故障相 / To fault *)
        _bFault := TRUE;                     (* 同步锁存 / Latch *)
        _eCause := E_DL_RtcCause.ePhaseBad;  (* 成因：非法相位 / Cause: illegal phase *)
END_CASE

(* —— 段 5：出口映射（bError/eState 同源，R191） —— *)
eBand := _eBandI;                            (* 档位出口单点映射 / Band outlet mapping *)
bError := _bFault;                           (* 故障标志镜像 / Fault flag mirror *)
eState := _eState;                           (* 状态出口 / State outlet *)
eCause := _eCause;                           (* 成因出口 / Cause outlet *)
END_FUNCTION_BLOCK

(* ---- FB_DL_RoPermeateQualityWatch.st ---- *)
(*
  Name: FB_DL_RoPermeateQualityWatch
  Category: DL_Process
  Version: 1.0.0
  Round: R90 / 2026-11-25
  开源溯源：clean-room 自研（族 RO/NF 膜法水处理，ST 开源生态实测 0 命中，无外部代码引入）
  功能：1) 产水电导率超限监视：越过上限后先经 tDebounceS 去抖（TON），去抖确认才置报警，
           避免单点尖峰造成误报警与误切段。
        2) 回差释放：报警锁存后必须回落到「上限 − 回差带宽」以下才解除，回差带宽由 fHystUsCm 给出，
           防止电导率在上限附近抖振导致报警继电器反复翻转。
        3) 连续超限计数 iOverCnt 记录本次越限持续的扫描拍数，作为劣化速率的粗观测量；
           趋势方向 xRising 由本次采样与上一拍快照的差值给出，差值超过 DL_TREND_EPS 才判上升，
           防止末位噪声被当作趋势。
  边界条件：1) 非有限值闸：三路实值入参统一过 NOT(x > -DL_BIG AND x < DL_BIG)，
           同时拦 NaN 与 Inf；命中时报警与趋势均强制 FALSE 并回待机相。原因是 NaN 与任何数比较
           均为假，会让回差释放判据静默失效（报警永不释放），故必须前置拦截（R19）。
        2) 组态零闸：fLimitUsCm 必须 > DL_EPS、fHystUsCm 必须 >= 0 且 <= fLimitUsCm，
           否则回差下沿会落到负值，释放判据永不成立（死锁），故判组态无效并暂停监视。
        3) 回差下沿钳制：fLimitUsCm − fHystUsCm 结果再钳到 >= 0，防组态越界后下沿为负。
        4) 时间零闸：tDebounceS <= T#0S 时 TON 立即置 Q，等价于「无去抖、即时报警」；
           这是合法组态，不判无效，但语义在此声明，禁止下游按「必有延时」假设时序。
        5) 状态机兜底：CASE 全态覆盖 + ELSE 强制回故障相；故障解除路径为 xEn 下降沿（可达）。
        6) FB 主体不使用 RETURN（跨平台可移植性考虑，统一单出口）。
  量纲自证：fCondUsCm、fLimitUsCm、fHystUsCm 三者同为电导率 [uS/cm]，比较与相减量纲一致；
           回差下沿 = (uS/cm) − (uS/cm) = uS/cm；tDebounceS 为 [TIME]，与 TON 的 PT 同量纲；
           趋势差值 = (uS/cm) − (uS/cm) = uS/cm，与 DL_TREND_EPS 同量纲，未跨量纲相加。
  码表 Error codes（本件格 0090_02xx）:
    16#0090_0201 信息级：输入非有限或组态越界，监视暂停（不置故障位，不阻止恢复）
    16#0090_0202 故障级：状态机落 ELSE 兜底（非法相位 ID），锁存至 xEn 下降沿解除
*)

TYPE E_DL_RpqwState :
(
    eRpqwIdle     := 0,    // 待机：未使能或输入无效 / Idle: disabled or invalid input
    eRpqwNormal   := 10,   // 正常：电导率在限值以下 / Normal: below limit
    eRpqwDebounce := 20,   // 去抖中：已越限，等待延时确认 / Debouncing: over limit, awaiting confirmation
    eRpqwAlarm    := 30,   // 报警：去抖确认后保持 / Alarm: confirmed and held
    eRpqwFault    := 90    // 故障：非法相位兜底 / Fault: illegal-phase fallback
);
END_TYPE

FUNCTION_BLOCK FB_DL_RoPermeateQualityWatch
VAR_INPUT
    xEn          : BOOL;    // 监视使能 [bool] / Monitoring enable [bool]
    fCondUsCm    : REAL;    // 产水电导率实测值 [uS/cm] / Permeate conductivity [uS/cm]
    fLimitUsCm   : REAL;    // 电导率报警上限 [uS/cm] / Conductivity alarm limit [uS/cm]
    fHystUsCm    : REAL;    // 报警释放回差带宽 [uS/cm] / Alarm release hysteresis band [uS/cm]
    tDebounceS   : TIME;    // 超限去抖延时 [TIME] / Over-limit debounce time [TIME]
END_VAR
VAR_OUTPUT
    xAlarm       : BOOL;    // 超限报警（带回差释放）[bool] / Over-limit alarm with hysteresis [bool]
    xRising      : BOOL;    // 电导率趋势上升标志 [bool] / Rising conductivity trend flag [bool]
    xValid       : BOOL;    // 输入有效标志 [bool] / Input valid flag [bool]
    iOverCnt     : INT;     // 连续超限扫描拍计数 [-] / Consecutive over-limit cycle count [-]
    eState       : E_DL_RpqwState;   // 状态出口，段尾单点映射 / State outlet, single-point mapped
    nErrId       : UDINT;   // 事件码，0 = 无事件 / Event code, 0 = none
END_VAR
VAR
    tonDeb       : TON;     // 超限去抖定时器，每拍无条件调用 / Debounce timer, unconditional call
    _eState      : E_DL_RpqwState := E_DL_RpqwState.eRpqwIdle;   // 内部相位（CASE 唯一写入目标）
    _fHystLoUsCm : REAL;    // 回差释放下沿 [uS/cm] / Hysteresis release low edge [uS/cm]
    _fCondPrev   : REAL;    // 上一拍电导率快照 [uS/cm] / Previous-cycle conductivity snapshot [uS/cm]
    _bOverUp     : BOOL;    // 越过上限（含触点）[bool] / Above upper limit, contact inclusive [bool]
    _bUnderDn    : BOOL;    // 回落到回差下沿以下 [bool] / Below hysteresis low edge [bool]
    _bCfgOk      : BOOL;    // 组态合法性聚合 [bool] / Configuration validity aggregate [bool]
    _bFault      : BOOL;    // 非法相位锁存位 [bool] / Illegal-phase latched flag [bool]
    _uInfo       : UDINT;   // 信息码，每拍重算 / Info code, recomputed every cycle
    _uFault      : UDINT;   // 故障码锁存 / Latched fault code
    _iOverCnt    : INT;     // 连续超限计数内部量 [-] / Consecutive over-limit internal counter [-]
END_VAR
VAR CONSTANT
    DL_EPS       : REAL := 1.0E-9;    // 组态零闸阈值 [-] / Configuration zero gate threshold [-]
    DL_BIG       : REAL := 1.0E12;    // 非有限值闸量级上限 [-] / Finiteness gate magnitude [-]
    DL_TREND_EPS : REAL := 0.05;      // 趋势判定的最小差值 [uS/cm] / Minimum delta for trend [uS/cm]
    DL_CNT_MAX   : INT  := 30000;     // 连续超限计数饱和上限 [-] / Over-limit counter saturation [-]
END_VAR

(* —— 段 1：单拍量预清零（锁存量 _uFault/_bFault/_iOverCnt/_fCondPrev 不入清单，R187①） —— *)
_uInfo := 16#0000_0000;                             // 信息码每拍重算 / Info code recomputed
nErrId := 16#0000_0000;                             // 事件码缺省无事件 / Event code defaults to none

(* —— 段 2：非有限值闸（R19：闸断比较通路，NaN 会让回差释放判据静默失效） —— *)
xValid := (fCondUsCm > -DL_BIG AND fCondUsCm < DL_BIG)          // 实测值有限
          AND (fLimitUsCm > -DL_BIG AND fLimitUsCm < DL_BIG)    // 限值有限
          AND (fHystUsCm > -DL_BIG AND fHystUsCm < DL_BIG);     // 回差带宽有限

(* —— 段 3：组态零闸与判据量（R4：回差下沿为负会使释放判据永不成立） —— *)
_bCfgOk := (fLimitUsCm > DL_EPS) AND (fHystUsCm >= 0.0) AND (fHystUsCm <= fLimitUsCm);
_fHystLoUsCm := MAX(0.0, fLimitUsCm - fHystUsCm);               // 回差下沿钳 >= 0 [uS/cm]
_bOverUp := _bCfgOk AND (fCondUsCm >= fLimitUsCm);              // 越过上限（含触点）
_bUnderDn := (NOT _bCfgOk) OR (fCondUsCm <= _fHystLoUsCm);      // 回落到下沿以下（组态坏视为释放）

(* —— 段 4：定时器无条件周期刷新（R7：调用语句不得置于 IF/CASE 内） —— *)
tonDeb(IN := xEn AND _bOverUp, PT := tDebounceS);   // 去抖窗，表达式入参，每拍必调

(* —— 段 5：相位机（只做迁移，出口在段 7 单点映射） —— *)
IF xValid THEN
    CASE _eState OF

    E_DL_RpqwState.eRpqwIdle:
        IF NOT xEn THEN
            ;                                       // 保持待机 / Stay idle
        ELSIF NOT _bCfgOk THEN
            _uInfo := 16#0090_0201;                 // 信息级：组态越界，暂停监视
        ELSIF _bOverUp AND tonDeb.Q THEN
            _eState := E_DL_RpqwState.eRpqwAlarm;   // 冷启动即在限上且已确认：直接报警
        ELSIF _bOverUp THEN
            _eState := E_DL_RpqwState.eRpqwDebounce;   // 越限但未确认：进去抖相
        ELSE
            _eState := E_DL_RpqwState.eRpqwNormal;  // 限下：进正常相
        END_IF

    E_DL_RpqwState.eRpqwNormal:
        IF (NOT xEn) OR (NOT _bCfgOk) THEN
            _eState := E_DL_RpqwState.eRpqwIdle;    // 失能或组态坏：退待机重判
        ELSIF _bOverUp THEN
            _eState := E_DL_RpqwState.eRpqwDebounce;   // 越过上限：进去抖相
        END_IF

    E_DL_RpqwState.eRpqwDebounce:
        IF NOT xEn THEN
            _eState := E_DL_RpqwState.eRpqwIdle;    // 失能即回待机
        ELSIF NOT _bOverUp THEN
            _eState := E_DL_RpqwState.eRpqwNormal;  // 去抖期间回落：撤销，回正常相
        ELSIF tonDeb.Q THEN
            _eState := E_DL_RpqwState.eRpqwAlarm;   // 去抖确认：报警锁存
        END_IF

    E_DL_RpqwState.eRpqwAlarm:
        IF NOT xEn THEN
            _eState := E_DL_RpqwState.eRpqwIdle;    // 失能清除报警
        ELSIF _bUnderDn THEN
            _eState := E_DL_RpqwState.eRpqwNormal;  // 回差释放：回正常相
        END_IF

    E_DL_RpqwState.eRpqwFault:
        IF NOT xEn THEN
            _bFault := FALSE;                       // 解除路径：xEn 下降沿（可达）
            _uFault := 16#0000_0000;
            _eState := E_DL_RpqwState.eRpqwIdle;
        END_IF

    ELSE
        _uFault := 16#0090_0202;                    // 故障级：非法相位 ID 兜底
        _bFault := TRUE;                            // 锁存（3 行内置，R45 配对）
        _eState := E_DL_RpqwState.eRpqwFault;       // 强制回故障相

    END_CASE

    (* —— 段 6：后置段（R23：计数一律在迁移判断之后处理） —— *)
    IF (_eState = E_DL_RpqwState.eRpqwNormal) OR (_eState = E_DL_RpqwState.eRpqwDebounce)
       OR (_eState = E_DL_RpqwState.eRpqwAlarm) THEN
        IF _bOverUp THEN
            _iOverCnt := MIN(DL_CNT_MAX, _iOverCnt + 1);   // 超限拍数累加（饱和）
        ELSE
            _iOverCnt := 0;                                 // 回落即清零
        END_IF
    ELSE
        _iOverCnt := 0;                                     // 非监视相一律清零
    END_IF
ELSE
    xAlarm := FALSE;                                // 报警强制 FALSE，无效数据不报警
    xRising := FALSE;                               // 趋势强制 FALSE
    _uInfo := 16#0090_0201;                         // 信息级：监视暂停
    _eState := E_DL_RpqwState.eRpqwIdle;            // 回待机相，等输入恢复
    _iOverCnt := 0;                                 // 计数清零（无效数据不累积）
END_IF

(* —— 段 7：出口单点映射（名实同源；报警由状态导出，不在多分支各写一遍） —— *)
xAlarm := (_eState = E_DL_RpqwState.eRpqwAlarm) AND (NOT _bFault);          // 报警出口
xRising := ((fCondUsCm - _fCondPrev) > DL_TREND_EPS) AND xValid AND (NOT _bFault);   // 趋势出口
iOverCnt := _iOverCnt;                              // 连续超限拍数出口
eState := _eState;                                  // 状态出口单点映射
IF _bFault THEN
    nErrId := _uFault;                              // 故障锁存码回放（禁同拍抹除）
ELSE
    nErrId := _uInfo;                               // 信息码
END_IF
_fCondPrev := fCondUsCm;                            // 快照统一在周期末尾更新（R23）

END_FUNCTION_BLOCK

(* ---- FB_DL_RotaryIndexModulo.st ---- *)
// =====================================================================
// FB_DL_RotaryIndexModulo.st
// 转盘工位索引与入料放行联锁（显式回绕禁 MOD+1、到位去抖 2 拍）
// Rotary table index and entry permit interlock FB
// 码位: 16#0005_045D ~ 16#0005_0461 (本件独占 5 槽)
// 修改记录: R29 初版 (按 DISPATCH_R29 序 19)
// =====================================================================
FUNCTION_BLOCK FB_DL_RotaryIndexModulo
VAR_INPUT
    bEnable      : BOOL  := FALSE;    // 使能 / Enable
    bIndexReq    : BOOL  := FALSE;    // 分度请求（上升沿受理）/ Index request on edge
    bReset       : BOOL  := FALSE;    // 复位 / Reset
    bAtPos       : BOOL  := FALSE;    // 转盘到位信号 / At position
    bIndexDone   : BOOL  := FALSE;    // 分度电机完成 / Index done
    bEntryClear  : BOOL  := FALSE;    // 入料通道已清空 / Entry clear
    uStationCnt  : USINT  := 8;       // 工位数 1~64 / Station count
    uStationInit : USINT  := 1;       // 初始工位号 1~64 / Initial station
    tIndexMax    : TIME  := T#5S;     // 分度超时 T#200MS~T#60S / Index timeout [s]
END_VAR
VAR_OUTPUT
    uStationIdx  : USINT;             // 当前工位号 1~64 / Station index
    bPermitEntry : BOOL;              // 入料放行 / Entry permit
    bIndexing    : BOOL;              // 分度中 / Indexing
    uIndexCnt    : UDINT;             // 累计分度次数 / Index count
    eErr         : UDINT;             // 错误码 / Error code
END_VAR
VAR
    rtrigReq     : R_TRIG;            // 分度请求沿检测（无条件刷新）/ Request edge detector
    tonIndex     : TON;               // 分度超时定时器（无条件刷新）/ Index timeout timer
    uAtPosDeb    : USINT;             // 到位去抖计数（连续 2 拍稳定）/ At-position debounce counter
    bAtPosStable : BOOL;              // 去抖后到位 / Stable at-position
    bTimeoutLatch: BOOL := FALSE;     // 超时锁存 / Timeout latch
    tIndexMaxS   : REAL;              // 超时秒值 / Timeout seconds [s]
    xFirstScan   : BOOL  := TRUE;     // 首扫标记 / First-scan flag
END_VAR

// ---------------------------------------------------------------------
// 代码位表（本件独占，勿复用）:
//   16#0005_045D 信息 正常（等待分度 / 已放行）
//   16#0005_045E 故障 tIndexMax 非法
//   16#0005_045F 故障 uStationCnt = 0 / uStationInit > uStationCnt（组态错）
//   16#0005_0460 信息 分度被拒（bEntryClear=FALSE 或 bAtPos=FALSE）→ bPermitEntry 保持 TRUE
//   16#0005_0461 故障 分度超 tIndexMax 未到位 → 关闭入料并锁存；解除=bReset 且 bAtPos 且 bEntryClear
// ---------------------------------------------------------------------

// ---- 超时秒值 / Timeout seconds ----
tIndexMaxS := TIME_TO_REAL(tIndexMax) / 1000.0;     // 秒值 / Seconds [s]

// ---- 请求沿检测（无条件刷新）/ Request edge, unconditional ----
rtrigReq(CLK := bIndexReq);     // 沿检测 / Edge detection

// ---- 超时参数闸 / Timeout validity gate ----
IF (tIndexMax = T#0MS) OR (tIndexMaxS < 0.2) OR (tIndexMaxS > 60.0) THEN
    bPermitEntry := FALSE;      // 放行撤销（安全侧）/ Permit off
    bIndexing := FALSE;         // 非分度 / Not indexing
    eErr := 16#0005_045E;       // 故障码 / Fault code
    RETURN;                     // 本拍结束 / End of cycle
END_IF

// ---- 组态错闸 / Configuration fault gate ----
IF (uStationCnt = 0) OR (uStationInit > uStationCnt) THEN
    bPermitEntry := FALSE;      // 放行撤销 / Permit off
    bIndexing := FALSE;         // 非分度 / Not indexing
    uStationIdx := 0;           // 工位号失效 / Index invalid
    eErr := 16#0005_045F;       // 故障码 / Fault code
    RETURN;                     // 本拍结束 / End of cycle
END_IF

// ---- 首扫初始化（R16 首扫纪律：bPermitEntry=FALSE 等首次到位确认）/ First-scan init ----
IF xFirstScan THEN
    uStationIdx := uStationInit;    // 初始工位号 / Init station
    bPermitEntry := FALSE;      // 首扫不放行 / No release on first scan
    bIndexing := FALSE;         // 非分度 / Not indexing
    xFirstScan := FALSE;        // 清标记 / Clear flag
END_IF

// ---- 使能撤销 / Disable ----
IF NOT bEnable THEN
    bPermitEntry := FALSE;      // 放行撤销 / Permit off
    bIndexing := FALSE;         // 非分度 / Not indexing
    bTimeoutLatch := FALSE;     // 锁存复位 / Latch reset
    eErr := 16#0005_045D;       // 信息级：空闲 / Info: idle
    RETURN;                     // 本拍结束 / End of cycle
END_IF

// ---- 超时锁存路径（解除 = bReset 且 bAtPos 且 bEntryClear）/ Timeout latch path ----
IF bTimeoutLatch THEN
    bPermitEntry := FALSE;      // 绝不带转盘运转放料 / Never release while latched
    bIndexing := FALSE;         // 非分度 / Not indexing
    eErr := 16#0005_0461;       // 故障码回放 / Fault code replay
    IF bReset AND bAtPos AND bEntryClear THEN
        bTimeoutLatch := FALSE;     // 解除锁存 / Release latch
        bPermitEntry := TRUE;       // 恢复放行 / Restore permit
        eErr := 16#0005_045D;       // 信息级：恢复 / Info: restored
    END_IF
    RETURN;                     // 本拍结束 / End of cycle
END_IF

// ---- 到位去抖（连续 2 拍稳定才认到位，防抖动）/ At-position debounce, 2 cycles ----
IF bAtPos THEN
    IF uAtPosDeb < 2 THEN
        uAtPosDeb := uAtPosDeb + 1;     // 稳定计数 / Stability count
    END_IF
ELSE
    uAtPosDeb := 0;             // 抖动复位 / Jitter reset
END_IF
bAtPosStable := (uAtPosDeb >= 2);   // 稳定到位 / Stable

// ---- 分度进行路径 / Indexing active path ----
IF bIndexing THEN
    tonIndex(IN := TRUE, PT := tIndexMax);  // 无条件刷新 / Unconditional refresh
    IF tonIndex.Q THEN
        // 分度超时未到位：关入料 + 锁存 / Timeout: close entry, latch
        bTimeoutLatch := TRUE;  // 锁存 / Latch
        bIndexing := FALSE;     // 非分度 / Not indexing
        bPermitEntry := FALSE;  // 关闭入料 / Close entry
        eErr := 16#0005_0461;   // 故障码 / Fault code
        RETURN;                 // 本拍结束 / End of cycle
    END_IF
    IF bIndexDone AND bAtPosStable THEN
        // 到位确认：工位号显式回绕（禁 MOD+1，防整除点出 0 工位）/ Explicit wrap, no MOD
        uStationIdx := uStationIdx + 1;     // 递增 / Increment
        IF uStationIdx > uStationCnt THEN
            uStationIdx := 1;   // 回绕到 1 / Wrap to 1
        END_IF
        uIndexCnt := uIndexCnt + 1;     // 累计分度 / Count
        bIndexing := FALSE;     // 分度结束 / Indexing off
        bPermitEntry := TRUE;   // 放行 / Release
        eErr := 16#0005_045D;   // 信息级：已放行 / Info: released
    END_IF
ELSE
    tonIndex(IN := FALSE, PT := tIndexMax);     // 定时器复位 / Timer reset

    // ---- 等待态：受理分度请求沿 / Waiting: accept request edge ----
    IF rtrigReq.Q AND bAtPosStable THEN
        IF bEntryClear THEN
            // 放行一次分度：先关入料 / Permit one index: close entry first
            bPermitEntry := FALSE;  // 关闭入料 / Close entry
            bIndexing := TRUE;      // 分度中 / Indexing
            eErr := 16#0005_045D;   // 信息级：分度中 / Info: indexing
        ELSE
            // 入料未清：拒绝分度（不停机但拒动），保持放行不误关料 / Entry not clear: reject, keep permit
            eErr := 16#0005_0460;   // 信息级：分度被拒 / Info: rejected
        END_IF
    ELSIF rtrigReq.Q AND (NOT bAtPosStable) THEN
        // 不在位：拒绝分度，保持放行 / Not at position: reject, keep permit
        eErr := 16#0005_0460;   // 信息级：分度被拒 / Info: rejected
    ELSE
        // 空闲等待：正常码（首扫确认后可放行）/ Idle waiting
        IF (NOT bPermitEntry) AND bAtPosStable AND bEntryClear THEN
            bPermitEntry := TRUE;   // 首次到位确认后放行 / Release after first confirm
        END_IF
        eErr := 16#0005_045D;   // 信息级：正常 / Info: normal
    END_IF
END_IF

END_FUNCTION_BLOCK

(* ---- FB_DL_SafetyDoorAuditBank.st ---- *)
(*
  FB_DL_SafetyDoorAuditBank  —  化成柜多安全门审计汇总（开门次数/批次锁定） / Formation cabinet multi-door audit bank: open counts and batch lock
  分类 Category : DL_Process
  版本 Version  : 1.0.0
  来源 Source   : t2-8-isa182 — 安全联锁审计族深化（与 I_DL_SafetyDoor 单门接口分工：那件管单门状态，本件管多门汇总）
  溯源 Origin   : clean-room 实现，未复制任何源码行
  功能 Function : 1) 8 门固定阵列逐门开门沿计数：每门 R_TRIG 阵列无条件周期刷新，
                  沿触发总计数 uOpenTotal 与分门计数 auOpenCnt 递增；
                  2) 批次锁定审计：bBatchLock 激活期任一门开门 → 0379 违约锁存
                  （独立记录首出违约门号 nViolDoor，R190 归因唯一）；
                  3) 审计饱和保护：uOpenTotal 逼近 UDINT 上限 → 停止递增并 037A
                  饱和锁存（防回绕伪造审计记录，还原方向不饱和原则）；
                  4) 相位机：eIdle（未使能）→ eAudit（审计中）→ eFault；
                  5) 信息级三码：开门计数沿 / 批次锁定激活 / 审计复位完成；
                  6) 解除式全当拍量（R240 落地），逐 BOOL 标注见段 4。
  边界 Boundary : ① 组态闸：bAuditEn = FALSE 相不计数不判违（审计仅使能相承载）；
                  ② 饱和反证句：饱和场景（累计达上限）不可由任何现有输出组合观测
                  （bError/nErrId 均无对应位），故独立占 037A；
                  ③ ELSE 兜底归并 037B 组态码（码表声明）；
                  ④ 无 GVL 依赖：纯引脚输入输出，无外部变量引用，无物理 IO 地址。
  依赖 Depends  : Standard.library（R_TRIG）
  码表 Error codes（Process 段 0005，窗口 0379~037B / 04A1~04A3）:
    16#0005_0379 故障级：批次锁定期间开门违约锁存（首出门号入 nViolDoor），锁存至 bReset
    16#0005_037A 故障级：审计总计数饱和锁存（停止递增防回绕），锁存至 bReset
    16#0005_037B 故障级：相位落 ELSE 兜底（归并声明），锁存至 bReset
    16#0005_04A1 信息级：开门计数沿（任一门开门沿触发）
    16#0005_04A2 信息级：批次锁定激活沿（进锁定审计态）
    16#0005_04A3 信息级：审计计数复位完成沿（bCountRst 生效拍）
  修订历史 Revision :
    2026-11-19  v1.0.0  R42 首版（批次 1 · 序号 4）
*)

TYPE E_DL_SdaState :
(
    eIdle   := 0,    // 未使能：不计数不判违 / Idle, not counting
    eAudit  := 10,   // 审计中：开门沿计数与批次违例监视 / Audit, counting and lock watch
    eFault  := 90    // 故障：违约或饱和锁定 / Fault, latched
);
END_TYPE

FUNCTION_BLOCK FB_DL_SafetyDoorAuditBank
VAR_INPUT
    a_bDoorOpen  : ARRAY[0..7] OF BOOL;  // 8 门开门反馈阵列，TRUE = 开 [-] / Door-open feedback array
    bAuditEn     : BOOL := FALSE;        // 审计使能（电平）[-] / Audit enable, level
    bBatchLock   : BOOL := FALSE;        // 批次锁定（电平），锁定期开门即违例 [-] / Batch lock, level
    bCountRst    : BOOL := FALSE;        // 计数复位指令，上升沿清全部计数 [-] / Count reset command edge
    bReset       : BOOL := FALSE;        // 复位，上升沿清故障锁存 / Reset edge clears fault latch
END_VAR
VAR_OUTPUT
    eState       : E_DL_SdaState;     // 状态出口，段尾单点映射 / State outlet
    uOpenTotal   : UDINT;             // 开门总计数 [次]，饱和即锁 / Total open count
    auOpenCnt    : ARRAY[0..7] OF UDINT;  // 分门开门计数 [次] / Per-door open counts
    nViolDoor    : USINT;             // 首出违约门号 [0..7]，255 = 无违约 / First violating door index
    bError       : BOOL;              // 故障锁存标志 / Fault latch flag
    nErrId       : UDINT;             // 事件码，0 = 无事件 / Event code
END_VAR
VAR
    a_rtDoor     : ARRAY[0..7] OF R_TRIG; // 8 门开门沿实例阵列，无条件刷新 / Door edge instance array
    rtCountRst   : R_TRIG;            // 计数复位沿实例，无条件刷新 / Count reset edge instance
    rtReset      : R_TRIG;            // 复位沿实例，无条件刷新 / Reset edge instance
    _eState      : E_DL_SdaState := E_DL_SdaState.eIdle;  // 内部相位（CASE 唯一写入目标）/ Internal phase
    _bLockInfoSent: BOOL;             // 批次锁定信息沿单发标志 / Lock-info one-shot sent flag
    _nIdx        : DINT;              // 阵列循环索引 [-] / Array loop index
    _bAnyOpen    : BOOL;              // 任一门开当拍量 [-] / Any-door-open current-scan flag
    _bSatWarn    : BOOL;              // 饱和临近当拍量（距上限不足 8 次计数）[-] / Near-saturation flag
    _bFault      : BOOL;              // 故障锁存位（锁存量）/ Latched fault bit
    _uFault      : UDINT;             // 故障码锁存（锁存量）/ Latched fault code
    _uInfo       : UDINT;             // 信息码，每拍重算 / Transient info code
END_VAR

(* —— 段 0：沿实例无条件周期刷新（禁置于 IF/CASE 内） —— *)
_bAnyOpen := a_bDoorOpen[0] OR a_bDoorOpen[1] OR a_bDoorOpen[2] OR a_bDoorOpen[3]
          OR a_bDoorOpen[4] OR a_bDoorOpen[5] OR a_bDoorOpen[6] OR a_bDoorOpen[7];
                                        // 任一门开（当拍量，展开式判据）
FOR _nIdx := 0 TO 7 DO               // 8 门沿实例逐门刷新（每拍必调）
    a_rtDoor[_nIdx](CLK := a_bDoorOpen[_nIdx]);          // 开门沿（每拍必调）
END_FOR
_bSatWarn := (uOpenTotal >= 16#FFFFFFF8);            // 饱和临近（距上限不足 8 计数槽）
rtCountRst(CLK := bCountRst);                        // 计数复位沿（每拍必调）
rtReset(CLK := bReset);                              // 复位沿（每拍必调）

(* —— 段 1：单拍量预清零（锁存量 _bFault/_uFault 不入清单，禁同拍抹除） —— *)
_uInfo := 16#0000_0000;             // 信息码每拍重算
nErrId := 16#0000_0000;             // 事件码缺省无事件

(* —— 段 2：复位沿 + 计数复位沿（判据当拍量） —— *)
IF rtReset.Q THEN                   // rtReset.Q = 当拍量
    _bFault := FALSE;               // 清故障锁存位
    _uFault := 16#0000_0000;        // 清故障锁存码
    nViolDoor := 255;               // 违约门号恢复哨兵 255 = 无违约
END_IF
IF rtCountRst.Q AND (NOT _bAnyOpen) THEN             // 复位沿 + 全部关门（当拍量）才可清零
    uOpenTotal := 16#0000_0000;     // 总计数清零
    FOR _nIdx := 0 TO 7 DO          // 分门计数清零
        auOpenCnt[_nIdx] := 16#0000_0000;    // 逐门清零
    END_FOR
    _uInfo := 16#0005_04A3;         // 信息级：审计复位完成沿
END_IF

(* —— 段 3：开门沿计数与违约/饱和锁存（判据当拍量；每拍至多递增一次净额） —— *)
FOR _nIdx := 0 TO 7 DO              // 逐门开门沿审计（每门独立归因）
    IF a_rtDoor[_nIdx].Q AND (_eState = E_DL_SdaState.eAudit) THEN
        IF bBatchLock AND (NOT _bFault) AND (nViolDoor = 255) THEN
            _uFault := 16#0005_0379;        // 故障级：批次锁定开门违约（首出门号锁定）
            _bFault := TRUE;                // 故障标志与码位配对（R45）
            nViolDoor := USINT_TO_USINT(_nIdx);     // 首出违约门号（DINT 收窄，域 0..7 结构性安全）
        ELSIF NOT _bSatWarn THEN
            uOpenTotal := uOpenTotal + 1;   // 总计数递增（饱和临近期停止）
            auOpenCnt[_nIdx] := auOpenCnt[_nIdx] + 1;   // 分门计数递增
            _uInfo := 16#0005_04A1;         // 信息级：开门计数沿
        END_IF
    END_IF
END_FOR
IF _bSatWarn AND (_eState = E_DL_SdaState.eAudit) AND (NOT _bFault) THEN
    _uFault := 16#0005_037A;        // 故障级：审计总计数饱和锁存
    _bFault := TRUE;
END_IF

(* —— 段 4：故障解除式（R240 落地，逐 BOOL 标注）：
     rtReset.Q = 当拍量；NOT _bAnyOpen = 当拍量；NOT bBatchLock = 当拍量。
     均不含锁存量（_bFault/_uFault），解除边真实可达（关门 + 撤锁 + 复位沿）。 —— *)
IF rtReset.Q AND (NOT _bAnyOpen) AND (NOT bBatchLock) THEN
    _bFault := FALSE;               // 清故障锁存位（锁存量，仅此当拍量解除沿可清）
    _uFault := 16#0000_0000;        // 清故障锁存码（锁存量，仅本当拍量解除沿可清）
    IF _eState = E_DL_SdaState.eFault THEN
        _eState := E_DL_SdaState.eIdle;     // 故障相迁出：回未使能
    END_IF
END_IF

(* —— 段 5：相位机（CASE 全覆盖 + ELSE 兜底） —— *)
CASE _eState OF

E_DL_SdaState.eIdle:
    IF bAuditEn AND (NOT _bFault) THEN
        _eState := E_DL_SdaState.eAudit;    // 使能：进审计相
    END_IF

E_DL_SdaState.eAudit:
    IF bBatchLock AND (NOT _bLockInfoSent) THEN
        _uInfo := 16#0005_04A2;             // 信息级：批次锁定激活沿（单发）
        _bLockInfoSent := TRUE;             // 沿单发标志
    END_IF
    IF NOT bBatchLock THEN
        _bLockInfoSent := FALSE;            // 撤锁重置单发标志
    END_IF
    IF NOT bAuditEn THEN
        _eState := E_DL_SdaState.eIdle;     // 撤使能：回未使能相
    END_IF
    (* 违约/饱和迁出在段 3 承载 *)

E_DL_SdaState.eFault:
    ;                                       // 故障相：等解除沿（段 4 承载迁出）

ELSE
    _uFault := 16#0005_037B;                // 故障级：非法相位兜底
    _bFault := TRUE;
    _eState := E_DL_SdaState.eFault;        // 强制回故障相

END_CASE

(* —— 段 6：出口单点映射（名实同源；锁存码回放，禁同拍抹除） —— *)
IF _bFault THEN
    nErrId := _uFault;              // 故障锁存码回放
ELSE
    nErrId := _uInfo;               // 信息码
END_IF
bError := _bFault;                  // 故障标志与锁存位同源
eState := _eState;                  // 状态出口单点映射

END_FUNCTION_BLOCK
